// TIA Portal V17 export
// export: Created 2025-07-28T08:20:46.6725827Z, ExportSetting WithDefaults, DisplayName Totally Integrated Automation Portal, DisplayVersion V17, DisplayName TIA Portal Openness, DisplayVersion V17, DisplayName TIA Portal Version Control Interface, DisplayVersion V17, DisplayName SINAMICS Startdrive Advanced, DisplayVersion V17, DisplayName SINAMICS Startdrive G130, G150, S120, S150, SINAMICS MV, S210, DisplayVersion V17, DisplayName SINAMICS Startdrive G110M, G120, G120C, G120D, G120P, G115D, DisplayVersion V17, DisplayName STEP 7 Professional, DisplayVersion V17, DisplayName STEP 7 Safety, DisplayVersion V17, DisplayName WinCC Professional, DisplayVersion V17
FUNCTION_BLOCK "S31808022001_Sequence_All_73b5c5_cfdfd9eb-ebd8-4267-a68e-df0ebcea3fa8 - Copy (2)_f93786"   // FB1, LAD
VERSION : 0.1
// stored: AutoNumber true, IsIECCheckEnabled false, UDAEnableTagReadback false
   VAR_INPUT
      iAutoRunning : Bool;
      iFaultReset : Bool;
      iOTS_Frm_Prev_TTDown : Bool;
      iOTS_Frm_Prev_TTUp : Bool;
      iPalletNtPrsntAtTTDown : Bool;
      iPalletNtPrsntAtTTUp : Bool;
      iPalletPrsnt_TTDown : Bool;
      iPalletPrsnt_TTUp : Bool;
      iPartReject : Bool;
      iRTR_Frm_Next_0DegTTUp : Bool;
      iRTR_Frm_Next_90DegTTUp : Bool;
      iRTR_Frm_Next_TTDown : Bool;
      iRecvAreaClr_TTDown : Bool;
      iRecvAreaClr_TTUp : Bool;
      iReset_fault : Bool;
      iRx_Frm_Prev_TTUp : Bool;
      iSstMode : Bool;
      iSstPB : Bool;
      iStprRaise_TTDown : Bool;
      iStprRaise_TTUp : Bool;
      iTTAt0Pos : Bool;
      iTTAt90Pos : Bool;
      iTTLocked : Bool;
      iTTUnlocked : Bool;
      iXferAreaClr_0DegTTDown : Bool;
      iXferAreaClr_0DegTTUp : Bool;
      iXferAreaClr_90DegTTUp : Bool;
   END_VAR
   VAR_OUTPUT
      qConvRun_TTDown : Bool;
      qConvRun_TTUp : Bool;
      qDelStprDown_TTUp : Bool;
      qOTS_Frm_TTDown : Bool;
      qOTS_Frm_TTUp : Bool;
      qOutput1 : Bool;
      qProcessStart : Bool;
      qRTR_Frm_TTDwn : Bool;
      qRTR_Frm_TTUp : Bool;
      qStprDown_TTDown : Bool;
      qStprDown_TTUp : Bool;
      qStprRaise_TTDown : Bool;
      qStprRaise_TTUp : Bool;
      qTTLockCmd : Bool;
      qTTUnlockCmd : Bool;
      qTT_0Deg : Bool;
      qTT_90Deg : Bool;
   END_VAR
   VAR_IN_OUT
      iqRX_Frn_Prev_TtDown : Bool;
      iqRx_Frm_Prev_TTUp : Bool;
      iqTx_To_Next_0DegTTDown : Bool;
      iqTx_To_Next_0DegTTUp : Bool;
      iqTx_To_Next_90DegTTUp : Bool;
   END_VAR
   VAR DB_SPECIFIC
      StateNo : Int;
      s100_StWtForTTUnlck : Bool;
      s100_StWtForTTUnlck_T1 : Bool;
      s10_StRecoveryCondition : Bool;
      s10_StRecoveryCondition_T1 : Bool;
      s10_StRecoveryCondition_T2 : Bool;
      s10_StRecoveryCondition_T3 : Bool;
      s10_StRecoveryCondition_T4 : Bool;
      s10_StRecoveryCondition_T5 : Bool;
      s10_StRecoveryCondition_T6 : Bool;
      s10_StRecoveryCondition_T7 : Bool;
      s110_StWtForTTTurn90 : Bool;
      s110_StWtForTTTurn90_T1 : Bool;
      s120_StWtForTTLck : Bool;
      s120_StWtForTTLck_T1 : Bool;
      s130_StChkTTDwnRdyToRecv : Bool;
      s130_StChkTTDwnRdyToRecv_T1 : Bool;
      s130_StChkTTDwnRdyToRecv_T2 : Bool;
      s140_StWtFrConveyorStrt : Bool;
      s140_StWtFrConveyorStrt_T1 : Bool;
      s150_StChkNxtStRdyToRecvTTUp : Bool;
      s150_StChkNxtStRdyToRecvTTUp_T1 : Bool;
      s150_StChkNxtStRdyToRecvTTUp_T2 : Bool;
      s15_StWaitForManCorrection : Bool;
      s15_StWaitForManCorrection_T1 : Bool;
      s160_StWtFrStprDn_CnvyrStrt : Bool;
      s160_StWtFrStprDn_CnvyrStrt_T1 : Bool;
      s165_StWtPalAbsnt : Bool;
      s165_StWtPalAbsnt_T1 : Bool;
      s167_StWtFrDeforkOvr : Bool;
      s167_StWtFrDeforkOvr_Cond1 : Bool;
      s167_StWtFrDeforkOvr_Cond2 : Bool;
      s167_StWtFrDeforkOvr_T1 : Bool;
      s170_StWtForTTUpStprUp : Bool;
      s170_StWtForTTUpStprUp_T1 : Bool;
      s180_StWtForTTUnlk : Bool;
      s180_StWtForTTUnlk_T1 : Bool;
      s190_StWtForTT_To_0 : Bool;
      s190_StWtForTT_To_0_T1 : Bool;
      s192_StWtForTTlok : Bool;
      s192_StWtForTTlok_T1 : Bool;
      s20_StChkForPalletPresent : Bool;
      s20_StChkForPalletPresent_T1 : Bool;
      s20_StChkForPalletPresent_T2 : Bool;
      s20_StChkForPalletPresent_T3 : Bool;
      s20_StChkForPalletPresent_T4 : Bool;
      s210_StWtFrTTUnlk : Bool;
      s210_StWtFrTTUnlk_T1 : Bool;
      s220_StWtFrTT_Trn_0 : Bool;
      s220_StWtFrTT_Trn_0_T1 : Bool;
      s230_StWtFrTTLock : Bool;
      s230_StWtFrTTLock_T1 : Bool;
      s240_StWtFRTRNxtStnTTDown : Bool;
      s240_StWtFRTRNxtStnTTDown_T1 : Bool;
      s240_StWtFRTRNxtStnTTDown_T2 : Bool;
      s250_StWtTTDnStprDn_CnvyrStr : Bool;
      s250_StWtTTDnStprDn_CnvyrStr_T1 : Bool;
      s260_StWtPalAbsent : Bool;
      s260_StWtPalAbsent_T1 : Bool;
      s270_StWtFrTTDwnStprUp : Bool;
      s270_StWtFrTTDwnStprUp_T1 : Bool;
      s280_StWtRFrOTSFRmPrev_TTUp : Bool;
      s280_StWtRFrOTSFRmPrev_TTUp_T1 : Bool;
      s290_StWtFrTTUpCnvyrStrt : Bool;
      s290_StWtFrTTUpCnvyrStrt_T1 : Bool;
      s300_StChkTTPos : Bool;
      s300_StChkTTPos_T1 : Bool;
      s300_StChkTTPos_T2 : Bool;
      s300_StChkTTPos_T3 : Bool;
      s30_StChckPartSts : Bool;
      s30_StChckPartSts_T1 : Bool;
      s310_StWtRTRFrmTTUpAt0 : Bool;
      s310_StWtRTRFrmTTUpAt0_T1 : Bool;
      s310_StWtRTRFrmTTUpAt0_T2 : Bool;
      s320_StWtFrTTUpCnvyrStrtAt0 : Bool;
      s320_StWtFrTTUpCnvyrStrtAt0_T1 : Bool;
      s340_StChkTTDwnRdyToRecvAt90 : Bool;
      s340_StChkTTDwnRdyToRecvAt90_T1 : Bool;
      s340_StChkTTDwnRdyToRecvAt90_T2 : Bool;
      s350_StWtCnvyrStrt90 : Bool;
      s350_StWtCnvyrStrt90_T1 : Bool;
      s365_StWtForTTUlkAtIbtwn : Bool;
      s365_StWtForTTUlkAtIbtwn_T1 : Bool;
      s370_StWtForTTTurnZrAtIbtwn : Bool;
      s370_StWtForTTTurnZrAtIbtwn_T1 : Bool;
      s380_StWtForTTLock : Bool;
      s380_StWtForTTLock_T1 : Bool;
      s400_StWt2Defork : Bool;
      s400_StWt2Defork_Cond1 : Bool;
      s400_StWt2Defork_Cond2 : Bool;
      s400_StWt2Defork_T1 : Bool;
      s40_StWtForTTUnlock : Bool;
      s40_StWtForTTUnlock_T1 : Bool;
      s410_StWtForTTUlkAtIbtwn : Bool;
      s410_StWtForTTUlkAtIbtwn_T1 : Bool;
      s415_StWtForTTTurn90AtIbtwn : Bool;
      s415_StWtForTTTurn90AtIbtwn_T1 : Bool;
      s420_StWtForTTLock1 : Bool;
      s420_StWtForTTLock1_T1 : Bool;
      s50_StWtForTTTurn0 : Bool;
      s50_StWtForTTTurn0_T1 : Bool;
      s60_StWtForTTLock : Bool;
      s60_StWtForTTLock_T1 : Bool;
      s70_StWtOTSfrmTTUp : Bool;
      s70_StWtOTSfrmTTUp_T1 : Bool;
      s80_StWtTTUpStpDwnCnvrStrt : Bool;
      s80_StWtTTUpStpDwnCnvrStrt_T1 : Bool;
      s85_StWtPalPresntAtRej : Bool;
      s85_StWtPalPresntAtRej_T1 : Bool;
      s90_StWtTTUpStprUp : Bool;
      s90_StWtTTUpStprUp_T1 : Bool;
      sDefork1Done : Bool;
      sDefork2Done : Bool;
      sOTSFrmDwnTout : Bool;
      sOTSFrmUpTout : Bool;
      sPalOnStop_TTDown : Bool;
      sPalOnStop_TTUp_0Deg : Bool;
      sPalOnStop_TTUp_90Deg : Bool;
      sPalletAbsnDebTTUp : Bool;
      sPalletAbsntDebTTDown : Bool;
      sPalletAbsntDebTTUp : Bool;
      sPalletPrsntDebTTDown : Bool;
      sPalletPrsntDebTTUp : Bool;
      sRTRFrmUpTout : Bool;
      sSst : Bool;
      sSstPulse : Bool;
      sSstRise : Bool;
      sStWtResetRel : Bool;
      sStWtResetRel_T1 : Bool;
      sTTDwnSeqOver : Bool;
      sTTDwn_0Pos_TX_Time : Bool;
      sTTDwn_90Pos_RX_Time : Bool;
      sTTDwn_Timer_ON : Bool;
      sTTUpSeqOver : Bool;
      sTTUp_90Pos_TX_Time : Bool;
      sTTUp_Timer_ON : Bool;
      sTrBothPalletPresent : Bool;
   END_VAR
   VAR_TEMP
      tOne : Bool;
   END_VAR
   VAR_TEMP   // added for the SCL form of the ladder/FBD networks
      _w1 : Bool;
   END_VAR
BEGIN

REGION Network 1
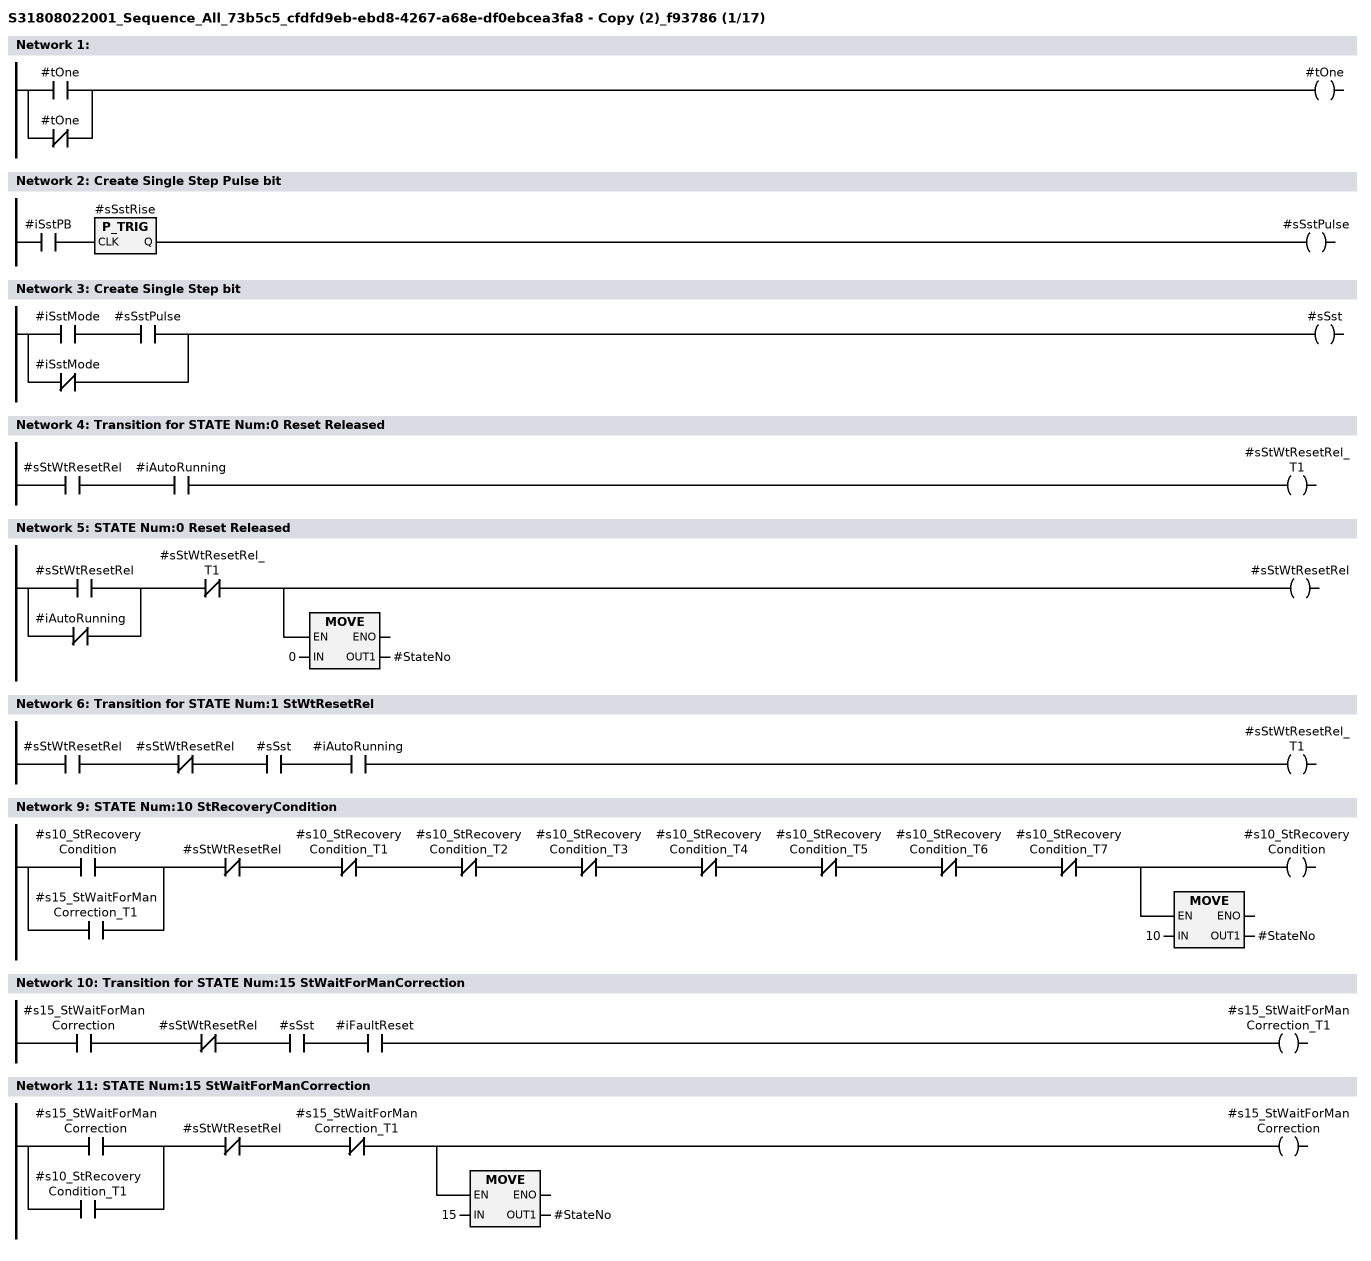
   RUNG wire#powerrail
      Contact( #tOne )
      wire#w1
      Coil( #tOne )
   END_RUNG
   RUNG wire#powerrail
      I_Contact( #tOne )
   END_RUNG wire#w1
   // the same network as SCL:
   #tOne := #tOne OR NOT #tOne;
END_REGION

REGION Network 2: Create Single Step Pulse bit
   RUNG wire#powerrail
      Contact( #iSstPB )
      P_Trig( #sSstRise )
      Coil( #sSstPulse )
   END_RUNG
   // the same network as SCL:
   #_w1 := #iSstPB AND NOT #sSstRise;   // rising edge
   #sSstRise := #iSstPB;
   #sSstPulse := #_w1;
END_REGION

REGION Network 3: Create Single Step bit
   RUNG wire#powerrail
      Contact( #iSstMode )
      Contact( #sSstPulse )
      wire#w1
      Coil( #sSst )
   END_RUNG
   RUNG wire#powerrail
      I_Contact( #iSstMode )
   END_RUNG wire#w1
   // the same network as SCL:
   #sSst := (#iSstMode AND #sSstPulse) OR NOT #iSstMode;
END_REGION

REGION Network 4: Transition for STATE Num:0 Reset Released
   RUNG wire#powerrail
      Contact( #sStWtResetRel )
      Contact( #iAutoRunning )
      Coil( #sStWtResetRel_T1 )
   END_RUNG
   // the same network as SCL:
   #sStWtResetRel_T1 := #sStWtResetRel AND #iAutoRunning;
END_REGION

REGION Network 5: STATE Num:0 Reset Released
   RUNG wire#powerrail
      Contact( #sStWtResetRel )
      wire#w1
      I_Contact( #sStWtResetRel_T1 )
      wire#w2
      Coil( #sStWtResetRel )
   END_RUNG
   RUNG wire#powerrail
      I_Contact( #iAutoRunning )
   END_RUNG wire#w1
   RUNG wire#w2
      { S7_GenerateENO := "TRUE" } Move(in := 0, out1 => #StateNo)
   END_RUNG
   // the same network as SCL:
   #sStWtResetRel := (#sStWtResetRel OR NOT #iAutoRunning) AND NOT #sStWtResetRel_T1;
   IF #sStWtResetRel THEN #StateNo := 0; END_IF;
END_REGION

REGION Network 6: Transition for STATE Num:1 StWtResetRel
   RUNG wire#powerrail
      Contact( #sStWtResetRel )
      I_Contact( #sStWtResetRel )
      Contact( #sSst )
      Contact( #iAutoRunning )
      Coil( #sStWtResetRel_T1 )
   END_RUNG
   // the same network as SCL:
   #sStWtResetRel_T1 := #sStWtResetRel AND NOT #sStWtResetRel AND #sSst AND #iAutoRunning;
END_REGION

NETWORK
TITLE = STATE Num:1 StWtResetRel
      A(;
      O     #sStWtResetRel;
//wrong transition variable removed
      );
      AN    #sStWtResetRel;
      AN    #sStWtResetRel_T1;
      =     %L1.0;
      A     %L1.0;
      BLD   102;
      =     #sStWtResetRel;
      A     %L1.0;
      JNB   Label_1;
      L     1;
      T     #StateNo;
Label_1:NOP   0;

NETWORK
TITLE = Transition for STATE Num:10 StRecoveryCondition
      A     #s10_StRecoveryCondition;
      AN    #sStWtResetRel;
      A     #sSst;
      =     %L1.0;
      A     %L1.0;
      A(;
      O(;
      A     #iRx_Frm_Prev_TTUp;
      AN    #iTTAt0Pos;
      );
      O(;
      A     #iqRX_Frn_Prev_TtDown;
      AN    #iTTAt90Pos;
      );
      O(;
      O     #iqTx_To_Next_90DegTTUp;
      O     #sPalOnStop_TTUp_90Deg;
      AN    #iTTAt90Pos;
      );
      O(;
      O     #iqTx_To_Next_0DegTTUp;
      O     #sPalOnStop_TTUp_0Deg;
      AN    #iTTAt0Pos;
      );
      O(;
      O     #iqTx_To_Next_0DegTTDown;
      O     #sPalOnStop_TTDown;
      AN    #iTTAt0Pos;
      );
      O(;
      O     #sPalOnStop_TTUp_0Deg;
      O     #sPalOnStop_TTUp_90Deg;
      O     #sPalOnStop_TTDown;
      A     #iTTUnlocked;
      );
      );
      =     #s10_StRecoveryCondition_T1;
      A     %L1.0;
      AN    #s10_StRecoveryCondition_T1;
      A(;
      O     #iqTx_To_Next_0DegTTUp;
      O     #sPalOnStop_TTUp_0Deg;
      );
      A     #iTTAt0Pos;
      A     #iTTLocked;
      =     #s10_StRecoveryCondition_T2;
      A     %L1.0;
      AN    #s10_StRecoveryCondition_T1;
      AN    #s10_StRecoveryCondition_T2;
      A(;
      O     #iqTx_To_Next_90DegTTUp;
      O     #sPalOnStop_TTUp_90Deg;
      );
      A     #iTTAt90Pos;
      A     #iTTLocked;
      =     #s10_StRecoveryCondition_T3;
      A     %L1.0;
      AN    #s10_StRecoveryCondition_T1;
      AN    #s10_StRecoveryCondition_T2;
      AN    #s10_StRecoveryCondition_T3;
      A(;
      O     #iqTx_To_Next_0DegTTDown;
      O     #sPalOnStop_TTDown;
      );
      A     #iTTAt0Pos;
      A     #iTTLocked;
      =     #s10_StRecoveryCondition_T4;
      A     %L1.0;
      AN    #s10_StRecoveryCondition_T1;
      AN    #s10_StRecoveryCondition_T2;
      AN    #s10_StRecoveryCondition_T3;
      AN    #s10_StRecoveryCondition_T4;
      A(;
      O     #iRx_Frm_Prev_TTUp;
      O     #iRecvAreaClr_TTUp;
      );
      A     #iTTAt0Pos;
      A     #iTTLocked;
      =     #s10_StRecoveryCondition_T5;
      A     %L1.0;
      AN    #s10_StRecoveryCondition_T1;
      AN    #s10_StRecoveryCondition_T2;
      AN    #s10_StRecoveryCondition_T3;
      AN    #s10_StRecoveryCondition_T4;
      AN    #s10_StRecoveryCondition_T5;
      A(;
      O     #iqRX_Frn_Prev_TtDown;
      ON    #iRecvAreaClr_TTDown;
      );
      A     #iTTAt90Pos;
      A     #iTTLocked;
      =     #s10_StRecoveryCondition_T6;
      A     %L1.0;
      AN    #s10_StRecoveryCondition_T1;
      AN    #s10_StRecoveryCondition_T2;
      AN    #s10_StRecoveryCondition_T3;
      AN    #s10_StRecoveryCondition_T4;
      AN    #s10_StRecoveryCondition_T5;
      AN    #s10_StRecoveryCondition_T6;
      A(;
      A(;
      A     #iXferAreaClr_90DegTTUp;
      A     #iXferAreaClr_0DegTTDown;
      A     #iRecvAreaClr_TTDown;
      A     #iRecvAreaClr_TTUp;
      );
      O(;
      AN    #sPalOnStop_TTUp_0Deg;
      AN    #sPalOnStop_TTUp_90Deg;
      AN    #sPalOnStop_TTDown;
      );
      O(;
      AN    #iqTx_To_Next_90DegTTUp;
      AN    #iqTx_To_Next_0DegTTUp;
      AN    #iqTx_To_Next_0DegTTDown;
      AN    #iqRX_Frn_Prev_TtDown;
      AN    #iRx_Frm_Prev_TTUp;
      );
      );
      =     #s10_StRecoveryCondition_T7;

REGION Network 9: STATE Num:10 StRecoveryCondition
   RUNG wire#powerrail
      Contact( #s10_StRecoveryCondition )
      wire#w1
      I_Contact( #sStWtResetRel )
      I_Contact( #s10_StRecoveryCondition_T1 )
      I_Contact( #s10_StRecoveryCondition_T2 )
      I_Contact( #s10_StRecoveryCondition_T3 )
      I_Contact( #s10_StRecoveryCondition_T4 )
      I_Contact( #s10_StRecoveryCondition_T5 )
      I_Contact( #s10_StRecoveryCondition_T6 )
      I_Contact( #s10_StRecoveryCondition_T7 )
      wire#w2
      Coil( #s10_StRecoveryCondition )
   END_RUNG
   RUNG wire#powerrail
      Contact( #s15_StWaitForManCorrection_T1 )
   END_RUNG wire#w1
   RUNG wire#w2
      { S7_GenerateENO := "TRUE" } Move(in := 10, out1 => #StateNo)
   END_RUNG
   // the same network as SCL:
   #s10_StRecoveryCondition := (#s10_StRecoveryCondition OR #s15_StWaitForManCorrection_T1) AND NOT #sStWtResetRel AND NOT #s10_StRecoveryCondition_T1 AND NOT #s10_StRecoveryCondition_T2 AND NOT #s10_StRecoveryCondition_T3 AND NOT #s10_StRecoveryCondition_T4 AND NOT #s10_StRecoveryCondition_T5 AND NOT #s10_StRecoveryCondition_T6 AND NOT #s10_StRecoveryCondition_T7;
   IF #s10_StRecoveryCondition THEN #StateNo := 10; END_IF;
END_REGION

REGION Network 10: Transition for STATE Num:15 StWaitForManCorrection
   RUNG wire#powerrail
      Contact( #s15_StWaitForManCorrection )
      I_Contact( #sStWtResetRel )
      Contact( #sSst )
      Contact( #iFaultReset )
      Coil( #s15_StWaitForManCorrection_T1 )
   END_RUNG
   // the same network as SCL:
   #s15_StWaitForManCorrection_T1 := #s15_StWaitForManCorrection AND NOT #sStWtResetRel AND #sSst AND #iFaultReset;
END_REGION

REGION Network 11: STATE Num:15 StWaitForManCorrection
   RUNG wire#powerrail
      Contact( #s15_StWaitForManCorrection )
      wire#w1
      I_Contact( #sStWtResetRel )
      I_Contact( #s15_StWaitForManCorrection_T1 )
      wire#w2
      Coil( #s15_StWaitForManCorrection )
   END_RUNG
   RUNG wire#powerrail
      Contact( #s10_StRecoveryCondition_T1 )
   END_RUNG wire#w1
   RUNG wire#w2
      { S7_GenerateENO := "TRUE" } Move(in := 15, out1 => #StateNo)
   END_RUNG
   // the same network as SCL:
   #s15_StWaitForManCorrection := (#s15_StWaitForManCorrection OR #s10_StRecoveryCondition_T1) AND NOT #sStWtResetRel AND NOT #s15_StWaitForManCorrection_T1;
   IF #s15_StWaitForManCorrection THEN #StateNo := 15; END_IF;
END_REGION

REGION Network 12: Transition for STATE Num:20 StChkForPalletPresent
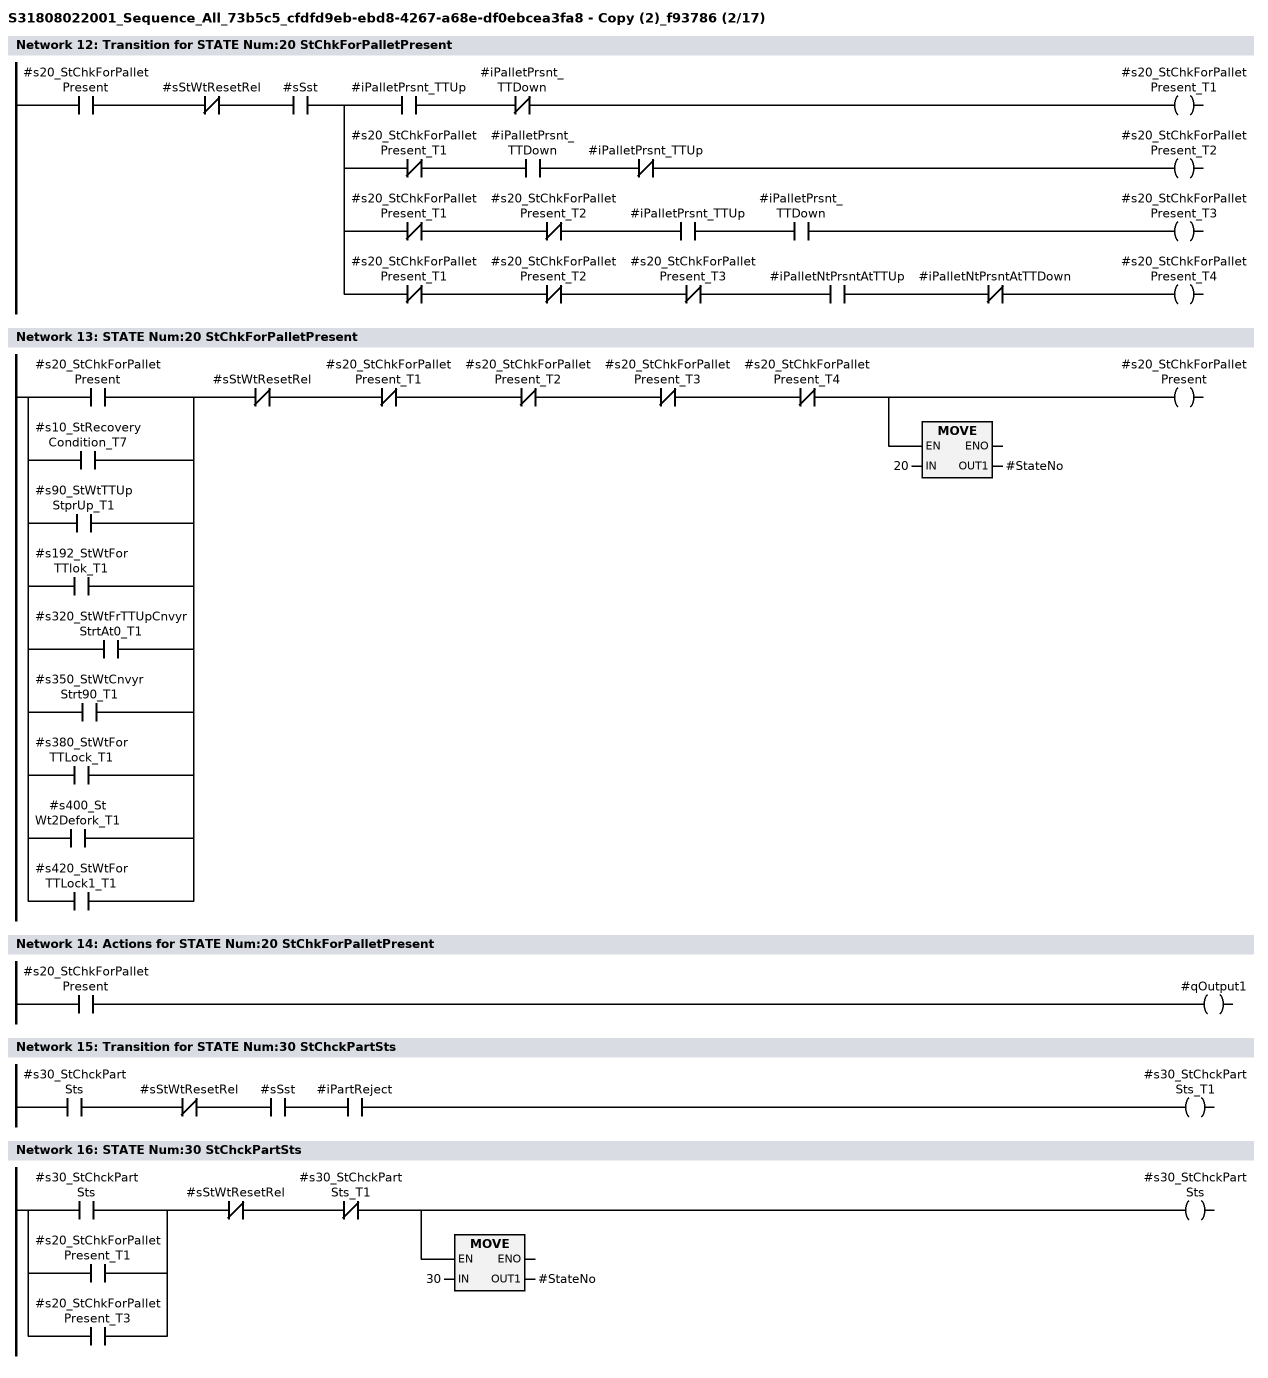
   RUNG wire#powerrail
      Contact( #s20_StChkForPalletPresent )
      I_Contact( #sStWtResetRel )
      Contact( #sSst )
      wire#w1
      Contact( #iPalletPrsnt_TTUp )
      I_Contact( #iPalletPrsnt_TTDown )
      Coil( #s20_StChkForPalletPresent_T1 )
   END_RUNG
   RUNG wire#w1
      I_Contact( #s20_StChkForPalletPresent_T1 )
      Contact( #iPalletPrsnt_TTDown )
      I_Contact( #iPalletPrsnt_TTUp )
      Coil( #s20_StChkForPalletPresent_T2 )
   END_RUNG
   RUNG wire#w1
      I_Contact( #s20_StChkForPalletPresent_T1 )
      I_Contact( #s20_StChkForPalletPresent_T2 )
      Contact( #iPalletPrsnt_TTUp )
      Contact( #iPalletPrsnt_TTDown )
      Coil( #s20_StChkForPalletPresent_T3 )
   END_RUNG
   RUNG wire#w1
      I_Contact( #s20_StChkForPalletPresent_T1 )
      I_Contact( #s20_StChkForPalletPresent_T2 )
      I_Contact( #s20_StChkForPalletPresent_T3 )
      Contact( #iPalletNtPrsntAtTTUp )
      I_Contact( #iPalletNtPrsntAtTTDown )
      Coil( #s20_StChkForPalletPresent_T4 )
   END_RUNG
   // the same network as SCL:
   #_w1 := #s20_StChkForPalletPresent AND NOT #sStWtResetRel AND #sSst;
   #s20_StChkForPalletPresent_T1 := #_w1 AND #iPalletPrsnt_TTUp AND NOT #iPalletPrsnt_TTDown;
   #s20_StChkForPalletPresent_T2 := #_w1 AND NOT #s20_StChkForPalletPresent_T1 AND #iPalletPrsnt_TTDown AND NOT #iPalletPrsnt_TTUp;
   #s20_StChkForPalletPresent_T3 := #_w1 AND NOT #s20_StChkForPalletPresent_T1 AND NOT #s20_StChkForPalletPresent_T2 AND #iPalletPrsnt_TTUp AND #iPalletPrsnt_TTDown;
   #s20_StChkForPalletPresent_T4 := #_w1 AND NOT #s20_StChkForPalletPresent_T1 AND NOT #s20_StChkForPalletPresent_T2 AND NOT #s20_StChkForPalletPresent_T3 AND #iPalletNtPrsntAtTTUp AND NOT #iPalletNtPrsntAtTTDown;
END_REGION

REGION Network 13: STATE Num:20 StChkForPalletPresent
   RUNG wire#powerrail
      Contact( #s20_StChkForPalletPresent )
      wire#w1
      I_Contact( #sStWtResetRel )
      I_Contact( #s20_StChkForPalletPresent_T1 )
      I_Contact( #s20_StChkForPalletPresent_T2 )
      I_Contact( #s20_StChkForPalletPresent_T3 )
      I_Contact( #s20_StChkForPalletPresent_T4 )
      wire#w2
      Coil( #s20_StChkForPalletPresent )
   END_RUNG
   RUNG wire#powerrail
      Contact( #s10_StRecoveryCondition_T7 )
   END_RUNG wire#w1
   RUNG wire#powerrail
      Contact( #s90_StWtTTUpStprUp_T1 )
   END_RUNG wire#w1
   RUNG wire#powerrail
      Contact( #s192_StWtForTTlok_T1 )
   END_RUNG wire#w1
   RUNG wire#powerrail
      Contact( #s320_StWtFrTTUpCnvyrStrtAt0_T1 )
   END_RUNG wire#w1
   RUNG wire#powerrail
      Contact( #s350_StWtCnvyrStrt90_T1 )
   END_RUNG wire#w1
   RUNG wire#powerrail
      Contact( #s380_StWtForTTLock_T1 )
   END_RUNG wire#w1
   RUNG wire#powerrail
      Contact( #s400_StWt2Defork_T1 )
   END_RUNG wire#w1
   RUNG wire#powerrail
      Contact( #s420_StWtForTTLock1_T1 )
   END_RUNG wire#w1
   RUNG wire#w2
      { S7_GenerateENO := "TRUE" } Move(in := 20, out1 => #StateNo)
   END_RUNG
   // the same network as SCL:
   #s20_StChkForPalletPresent := (#s20_StChkForPalletPresent OR #s10_StRecoveryCondition_T7 OR #s90_StWtTTUpStprUp_T1 OR #s192_StWtForTTlok_T1 OR #s320_StWtFrTTUpCnvyrStrtAt0_T1 OR #s350_StWtCnvyrStrt90_T1 OR #s380_StWtForTTLock_T1 OR #s400_StWt2Defork_T1 OR #s420_StWtForTTLock1_T1) AND NOT #sStWtResetRel AND NOT #s20_StChkForPalletPresent_T1 AND NOT #s20_StChkForPalletPresent_T2 AND NOT #s20_StChkForPalletPresent_T3 AND NOT #s20_StChkForPalletPresent_T4;
   IF #s20_StChkForPalletPresent THEN #StateNo := 20; END_IF;
END_REGION

REGION Network 14: Actions for STATE Num:20 StChkForPalletPresent
   RUNG wire#powerrail
      Contact( #s20_StChkForPalletPresent )
      Coil( #qOutput1 )
   END_RUNG
   // the same network as SCL:
   #qOutput1 := #s20_StChkForPalletPresent;
END_REGION

REGION Network 15: Transition for STATE Num:30 StChckPartSts
   RUNG wire#powerrail
      Contact( #s30_StChckPartSts )
      I_Contact( #sStWtResetRel )
      Contact( #sSst )
      Contact( #iPartReject )
      Coil( #s30_StChckPartSts_T1 )
   END_RUNG
   // the same network as SCL:
   #s30_StChckPartSts_T1 := #s30_StChckPartSts AND NOT #sStWtResetRel AND #sSst AND #iPartReject;
END_REGION

REGION Network 16: STATE Num:30 StChckPartSts
   RUNG wire#powerrail
      Contact( #s30_StChckPartSts )
      wire#w1
      I_Contact( #sStWtResetRel )
      I_Contact( #s30_StChckPartSts_T1 )
      wire#w2
      Coil( #s30_StChckPartSts )
   END_RUNG
   RUNG wire#powerrail
      Contact( #s20_StChkForPalletPresent_T1 )
   END_RUNG wire#w1
   RUNG wire#powerrail
      Contact( #s20_StChkForPalletPresent_T3 )
   END_RUNG wire#w1
   RUNG wire#w2
      { S7_GenerateENO := "TRUE" } Move(in := 30, out1 => #StateNo)
   END_RUNG
   // the same network as SCL:
   #s30_StChckPartSts := (#s30_StChckPartSts OR #s20_StChkForPalletPresent_T1 OR #s20_StChkForPalletPresent_T3) AND NOT #sStWtResetRel AND NOT #s30_StChckPartSts_T1;
   IF #s30_StChckPartSts THEN #StateNo := 30; END_IF;
END_REGION

REGION Network 17: Actions for STATE Num:30 StChckPartSts
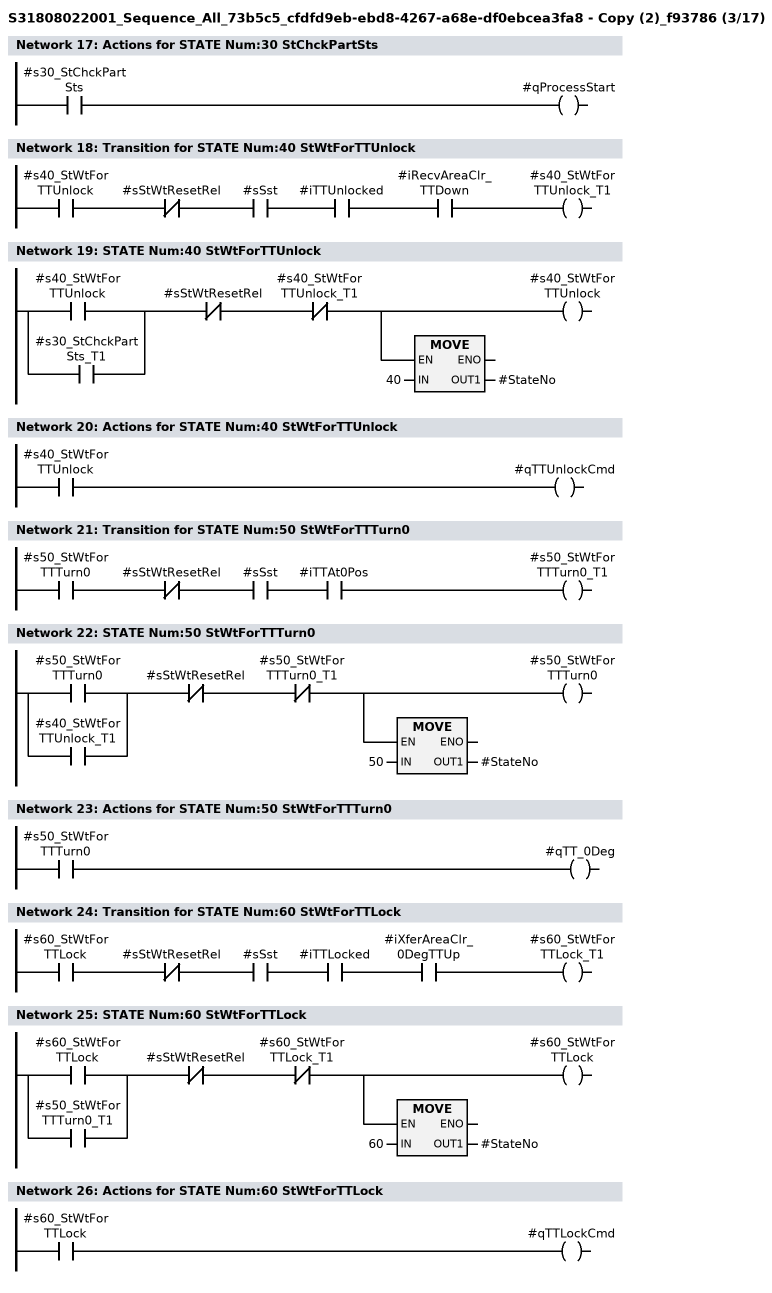
   RUNG wire#powerrail
      Contact( #s30_StChckPartSts )
      Coil( #qProcessStart )
   END_RUNG
   // the same network as SCL:
   #qProcessStart := #s30_StChckPartSts;
END_REGION

REGION Network 18: Transition for STATE Num:40 StWtForTTUnlock
   RUNG wire#powerrail
      Contact( #s40_StWtForTTUnlock )
      I_Contact( #sStWtResetRel )
      Contact( #sSst )
      Contact( #iTTUnlocked )
      Contact( #iRecvAreaClr_TTDown )
      Coil( #s40_StWtForTTUnlock_T1 )
   END_RUNG
   // the same network as SCL:
   #s40_StWtForTTUnlock_T1 := #s40_StWtForTTUnlock AND NOT #sStWtResetRel AND #sSst AND #iTTUnlocked AND #iRecvAreaClr_TTDown;
END_REGION

REGION Network 19: STATE Num:40 StWtForTTUnlock
   RUNG wire#powerrail
      Contact( #s40_StWtForTTUnlock )
      wire#w1
      I_Contact( #sStWtResetRel )
      I_Contact( #s40_StWtForTTUnlock_T1 )
      wire#w2
      Coil( #s40_StWtForTTUnlock )
   END_RUNG
   RUNG wire#powerrail
      Contact( #s30_StChckPartSts_T1 )
   END_RUNG wire#w1
   RUNG wire#w2
      { S7_GenerateENO := "TRUE" } Move(in := 40, out1 => #StateNo)
   END_RUNG
   // the same network as SCL:
   #s40_StWtForTTUnlock := (#s40_StWtForTTUnlock OR #s30_StChckPartSts_T1) AND NOT #sStWtResetRel AND NOT #s40_StWtForTTUnlock_T1;
   IF #s40_StWtForTTUnlock THEN #StateNo := 40; END_IF;
END_REGION

REGION Network 20: Actions for STATE Num:40 StWtForTTUnlock
   RUNG wire#powerrail
      Contact( #s40_StWtForTTUnlock )
      Coil( #qTTUnlockCmd )
   END_RUNG
   // the same network as SCL:
   #qTTUnlockCmd := #s40_StWtForTTUnlock;
END_REGION

REGION Network 21: Transition for STATE Num:50 StWtForTTTurn0
   RUNG wire#powerrail
      Contact( #s50_StWtForTTTurn0 )
      I_Contact( #sStWtResetRel )
      Contact( #sSst )
      Contact( #iTTAt0Pos )
      Coil( #s50_StWtForTTTurn0_T1 )
   END_RUNG
   // the same network as SCL:
   #s50_StWtForTTTurn0_T1 := #s50_StWtForTTTurn0 AND NOT #sStWtResetRel AND #sSst AND #iTTAt0Pos;
END_REGION

REGION Network 22: STATE Num:50 StWtForTTTurn0
   RUNG wire#powerrail
      Contact( #s50_StWtForTTTurn0 )
      wire#w1
      I_Contact( #sStWtResetRel )
      I_Contact( #s50_StWtForTTTurn0_T1 )
      wire#w2
      Coil( #s50_StWtForTTTurn0 )
   END_RUNG
   RUNG wire#powerrail
      Contact( #s40_StWtForTTUnlock_T1 )
   END_RUNG wire#w1
   RUNG wire#w2
      { S7_GenerateENO := "TRUE" } Move(in := 50, out1 => #StateNo)
   END_RUNG
   // the same network as SCL:
   #s50_StWtForTTTurn0 := (#s50_StWtForTTTurn0 OR #s40_StWtForTTUnlock_T1) AND NOT #sStWtResetRel AND NOT #s50_StWtForTTTurn0_T1;
   IF #s50_StWtForTTTurn0 THEN #StateNo := 50; END_IF;
END_REGION

REGION Network 23: Actions for STATE Num:50 StWtForTTTurn0
   RUNG wire#powerrail
      Contact( #s50_StWtForTTTurn0 )
      Coil( #qTT_0Deg )
   END_RUNG
   // the same network as SCL:
   #qTT_0Deg := #s50_StWtForTTTurn0;
END_REGION

REGION Network 24: Transition for STATE Num:60 StWtForTTLock
   RUNG wire#powerrail
      Contact( #s60_StWtForTTLock )
      I_Contact( #sStWtResetRel )
      Contact( #sSst )
      Contact( #iTTLocked )
      Contact( #iXferAreaClr_0DegTTUp )
      Coil( #s60_StWtForTTLock_T1 )
   END_RUNG
   // the same network as SCL:
   #s60_StWtForTTLock_T1 := #s60_StWtForTTLock AND NOT #sStWtResetRel AND #sSst AND #iTTLocked AND #iXferAreaClr_0DegTTUp;
END_REGION

REGION Network 25: STATE Num:60 StWtForTTLock
   RUNG wire#powerrail
      Contact( #s60_StWtForTTLock )
      wire#w1
      I_Contact( #sStWtResetRel )
      I_Contact( #s60_StWtForTTLock_T1 )
      wire#w2
      Coil( #s60_StWtForTTLock )
   END_RUNG
   RUNG wire#powerrail
      Contact( #s50_StWtForTTTurn0_T1 )
   END_RUNG wire#w1
   RUNG wire#w2
      { S7_GenerateENO := "TRUE" } Move(in := 60, out1 => #StateNo)
   END_RUNG
   // the same network as SCL:
   #s60_StWtForTTLock := (#s60_StWtForTTLock OR #s50_StWtForTTTurn0_T1) AND NOT #sStWtResetRel AND NOT #s60_StWtForTTLock_T1;
   IF #s60_StWtForTTLock THEN #StateNo := 60; END_IF;
END_REGION

REGION Network 26: Actions for STATE Num:60 StWtForTTLock
   RUNG wire#powerrail
      Contact( #s60_StWtForTTLock )
      Coil( #qTTLockCmd )
   END_RUNG
   // the same network as SCL:
   #qTTLockCmd := #s60_StWtForTTLock;
END_REGION

REGION Network 27: Transition for STATE Num:70 StWtOTSfrmTTUp
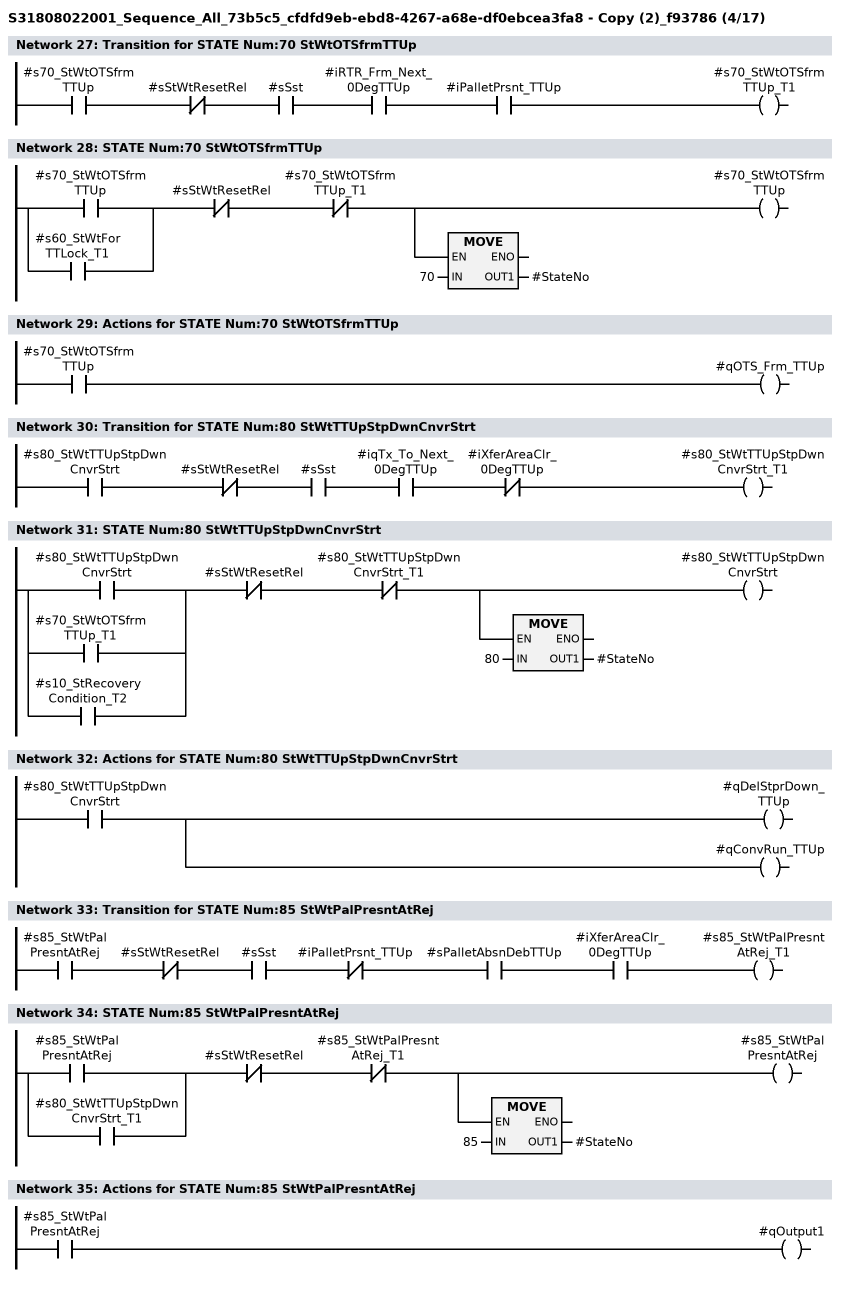
   RUNG wire#powerrail
      Contact( #s70_StWtOTSfrmTTUp )
      I_Contact( #sStWtResetRel )
      Contact( #sSst )
      Contact( #iRTR_Frm_Next_0DegTTUp )
      Contact( #iPalletPrsnt_TTUp )
      Coil( #s70_StWtOTSfrmTTUp_T1 )
   END_RUNG
   // the same network as SCL:
   #s70_StWtOTSfrmTTUp_T1 := #s70_StWtOTSfrmTTUp AND NOT #sStWtResetRel AND #sSst AND #iRTR_Frm_Next_0DegTTUp AND #iPalletPrsnt_TTUp;
END_REGION

REGION Network 28: STATE Num:70 StWtOTSfrmTTUp
   RUNG wire#powerrail
      Contact( #s70_StWtOTSfrmTTUp )
      wire#w1
      I_Contact( #sStWtResetRel )
      I_Contact( #s70_StWtOTSfrmTTUp_T1 )
      wire#w2
      Coil( #s70_StWtOTSfrmTTUp )
   END_RUNG
   RUNG wire#powerrail
      Contact( #s60_StWtForTTLock_T1 )
   END_RUNG wire#w1
   RUNG wire#w2
      { S7_GenerateENO := "TRUE" } Move(in := 70, out1 => #StateNo)
   END_RUNG
   // the same network as SCL:
   #s70_StWtOTSfrmTTUp := (#s70_StWtOTSfrmTTUp OR #s60_StWtForTTLock_T1) AND NOT #sStWtResetRel AND NOT #s70_StWtOTSfrmTTUp_T1;
   IF #s70_StWtOTSfrmTTUp THEN #StateNo := 70; END_IF;
END_REGION

REGION Network 29: Actions for STATE Num:70 StWtOTSfrmTTUp
   RUNG wire#powerrail
      Contact( #s70_StWtOTSfrmTTUp )
      Coil( #qOTS_Frm_TTUp )
   END_RUNG
   // the same network as SCL:
   #qOTS_Frm_TTUp := #s70_StWtOTSfrmTTUp;
END_REGION

REGION Network 30: Transition for STATE Num:80 StWtTTUpStpDwnCnvrStrt
   RUNG wire#powerrail
      Contact( #s80_StWtTTUpStpDwnCnvrStrt )
      I_Contact( #sStWtResetRel )
      Contact( #sSst )
      Contact( #iqTx_To_Next_0DegTTUp )
      I_Contact( #iXferAreaClr_0DegTTUp )
      Coil( #s80_StWtTTUpStpDwnCnvrStrt_T1 )
   END_RUNG
   // the same network as SCL:
   #s80_StWtTTUpStpDwnCnvrStrt_T1 := #s80_StWtTTUpStpDwnCnvrStrt AND NOT #sStWtResetRel AND #sSst AND #iqTx_To_Next_0DegTTUp AND NOT #iXferAreaClr_0DegTTUp;
END_REGION

REGION Network 31: STATE Num:80 StWtTTUpStpDwnCnvrStrt
   RUNG wire#powerrail
      Contact( #s80_StWtTTUpStpDwnCnvrStrt )
      wire#w1
      I_Contact( #sStWtResetRel )
      I_Contact( #s80_StWtTTUpStpDwnCnvrStrt_T1 )
      wire#w2
      Coil( #s80_StWtTTUpStpDwnCnvrStrt )
   END_RUNG
   RUNG wire#powerrail
      Contact( #s70_StWtOTSfrmTTUp_T1 )
   END_RUNG wire#w1
   RUNG wire#powerrail
      Contact( #s10_StRecoveryCondition_T2 )
   END_RUNG wire#w1
   RUNG wire#w2
      { S7_GenerateENO := "TRUE" } Move(in := 80, out1 => #StateNo)
   END_RUNG
   // the same network as SCL:
   #s80_StWtTTUpStpDwnCnvrStrt := (#s80_StWtTTUpStpDwnCnvrStrt OR #s70_StWtOTSfrmTTUp_T1 OR #s10_StRecoveryCondition_T2) AND NOT #sStWtResetRel AND NOT #s80_StWtTTUpStpDwnCnvrStrt_T1;
   IF #s80_StWtTTUpStpDwnCnvrStrt THEN #StateNo := 80; END_IF;
END_REGION

REGION Network 32: Actions for STATE Num:80 StWtTTUpStpDwnCnvrStrt
   RUNG wire#powerrail
      Contact( #s80_StWtTTUpStpDwnCnvrStrt )
      wire#w1
      Coil( #qDelStprDown_TTUp )
   END_RUNG
   RUNG wire#w1
      Coil( #qConvRun_TTUp )
   END_RUNG
   // the same network as SCL:
   #qDelStprDown_TTUp := #s80_StWtTTUpStpDwnCnvrStrt;
   #qConvRun_TTUp := #s80_StWtTTUpStpDwnCnvrStrt;
END_REGION

REGION Network 33: Transition for STATE Num:85 StWtPalPresntAtRej
   RUNG wire#powerrail
      Contact( #s85_StWtPalPresntAtRej )
      I_Contact( #sStWtResetRel )
      Contact( #sSst )
      I_Contact( #iPalletPrsnt_TTUp )
      Contact( #sPalletAbsnDebTTUp )
      Contact( #iXferAreaClr_0DegTTUp )
      Coil( #s85_StWtPalPresntAtRej_T1 )
   END_RUNG
   // the same network as SCL:
   #s85_StWtPalPresntAtRej_T1 := #s85_StWtPalPresntAtRej AND NOT #sStWtResetRel AND #sSst AND NOT #iPalletPrsnt_TTUp AND #sPalletAbsnDebTTUp AND #iXferAreaClr_0DegTTUp;
END_REGION

REGION Network 34: STATE Num:85 StWtPalPresntAtRej
   RUNG wire#powerrail
      Contact( #s85_StWtPalPresntAtRej )
      wire#w1
      I_Contact( #sStWtResetRel )
      I_Contact( #s85_StWtPalPresntAtRej_T1 )
      wire#w2
      Coil( #s85_StWtPalPresntAtRej )
   END_RUNG
   RUNG wire#powerrail
      Contact( #s80_StWtTTUpStpDwnCnvrStrt_T1 )
   END_RUNG wire#w1
   RUNG wire#w2
      { S7_GenerateENO := "TRUE" } Move(in := 85, out1 => #StateNo)
   END_RUNG
   // the same network as SCL:
   #s85_StWtPalPresntAtRej := (#s85_StWtPalPresntAtRej OR #s80_StWtTTUpStpDwnCnvrStrt_T1) AND NOT #sStWtResetRel AND NOT #s85_StWtPalPresntAtRej_T1;
   IF #s85_StWtPalPresntAtRej THEN #StateNo := 85; END_IF;
END_REGION

REGION Network 35: Actions for STATE Num:85 StWtPalPresntAtRej
   RUNG wire#powerrail
      Contact( #s85_StWtPalPresntAtRej )
      Coil( #qOutput1 )
   END_RUNG
   // the same network as SCL:
   #qOutput1 := #s85_StWtPalPresntAtRej;
END_REGION

REGION Network 36: Transition for STATE Num:90 StWtTTUpStprUp
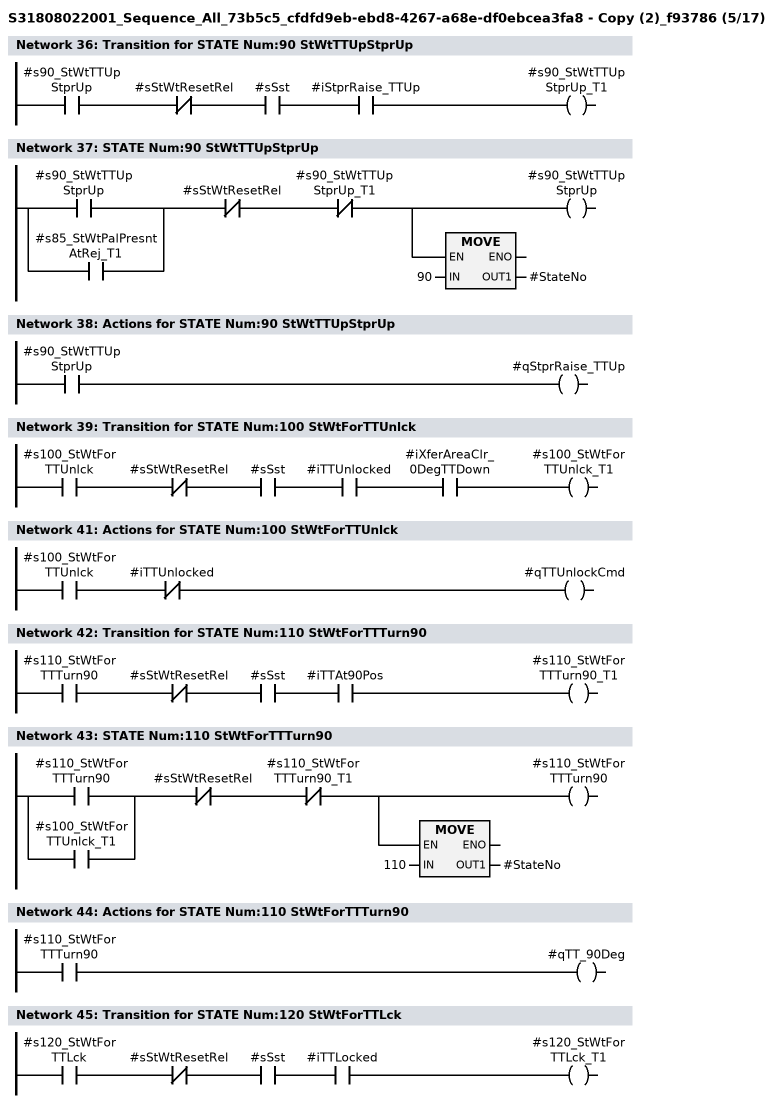
   RUNG wire#powerrail
      Contact( #s90_StWtTTUpStprUp )
      I_Contact( #sStWtResetRel )
      Contact( #sSst )
      Contact( #iStprRaise_TTUp )
      Coil( #s90_StWtTTUpStprUp_T1 )
   END_RUNG
   // the same network as SCL:
   #s90_StWtTTUpStprUp_T1 := #s90_StWtTTUpStprUp AND NOT #sStWtResetRel AND #sSst AND #iStprRaise_TTUp;
END_REGION

REGION Network 37: STATE Num:90 StWtTTUpStprUp
   RUNG wire#powerrail
      Contact( #s90_StWtTTUpStprUp )
      wire#w1
      I_Contact( #sStWtResetRel )
      I_Contact( #s90_StWtTTUpStprUp_T1 )
      wire#w2
      Coil( #s90_StWtTTUpStprUp )
   END_RUNG
   RUNG wire#powerrail
      Contact( #s85_StWtPalPresntAtRej_T1 )
   END_RUNG wire#w1
   RUNG wire#w2
      { S7_GenerateENO := "TRUE" } Move(in := 90, out1 => #StateNo)
   END_RUNG
   // the same network as SCL:
   #s90_StWtTTUpStprUp := (#s90_StWtTTUpStprUp OR #s85_StWtPalPresntAtRej_T1) AND NOT #sStWtResetRel AND NOT #s90_StWtTTUpStprUp_T1;
   IF #s90_StWtTTUpStprUp THEN #StateNo := 90; END_IF;
END_REGION

REGION Network 38: Actions for STATE Num:90 StWtTTUpStprUp
   RUNG wire#powerrail
      Contact( #s90_StWtTTUpStprUp )
      Coil( #qStprRaise_TTUp )
   END_RUNG
   // the same network as SCL:
   #qStprRaise_TTUp := #s90_StWtTTUpStprUp;
END_REGION

REGION Network 39: Transition for STATE Num:100 StWtForTTUnlck
   RUNG wire#powerrail
      Contact( #s100_StWtForTTUnlck )
      I_Contact( #sStWtResetRel )
      Contact( #sSst )
      Contact( #iTTUnlocked )
      Contact( #iXferAreaClr_0DegTTDown )
      Coil( #s100_StWtForTTUnlck_T1 )
   END_RUNG
   // the same network as SCL:
   #s100_StWtForTTUnlck_T1 := #s100_StWtForTTUnlck AND NOT #sStWtResetRel AND #sSst AND #iTTUnlocked AND #iXferAreaClr_0DegTTDown;
END_REGION

NETWORK
TITLE = STATE Num:100 StWtForTTUnlck
      A(;
      O     #s100_StWtForTTUnlck;
      );
      AN    #sStWtResetRel;
      AN    #s100_StWtForTTUnlck_T1;
      =     %L1.0;
      A     %L1.0;
      BLD   102;
      =     #s100_StWtForTTUnlck;
      A     %L1.0;
      JNB   Label_13;
      L     100;
      T     #StateNo;
Label_13:NOP   0;

REGION Network 41: Actions for STATE Num:100 StWtForTTUnlck
   RUNG wire#powerrail
      Contact( #s100_StWtForTTUnlck )
      I_Contact( #iTTUnlocked )
      Coil( #qTTUnlockCmd )
   END_RUNG
   // the same network as SCL:
   #qTTUnlockCmd := #s100_StWtForTTUnlck AND NOT #iTTUnlocked;
END_REGION

REGION Network 42: Transition for STATE Num:110 StWtForTTTurn90
   RUNG wire#powerrail
      Contact( #s110_StWtForTTTurn90 )
      I_Contact( #sStWtResetRel )
      Contact( #sSst )
      Contact( #iTTAt90Pos )
      Coil( #s110_StWtForTTTurn90_T1 )
   END_RUNG
   // the same network as SCL:
   #s110_StWtForTTTurn90_T1 := #s110_StWtForTTTurn90 AND NOT #sStWtResetRel AND #sSst AND #iTTAt90Pos;
END_REGION

REGION Network 43: STATE Num:110 StWtForTTTurn90
   RUNG wire#powerrail
      Contact( #s110_StWtForTTTurn90 )
      wire#w1
      I_Contact( #sStWtResetRel )
      I_Contact( #s110_StWtForTTTurn90_T1 )
      wire#w2
      Coil( #s110_StWtForTTTurn90 )
   END_RUNG
   RUNG wire#powerrail
      Contact( #s100_StWtForTTUnlck_T1 )
   END_RUNG wire#w1
   RUNG wire#w2
      { S7_GenerateENO := "TRUE" } Move(in := 110, out1 => #StateNo)
   END_RUNG
   // the same network as SCL:
   #s110_StWtForTTTurn90 := (#s110_StWtForTTTurn90 OR #s100_StWtForTTUnlck_T1) AND NOT #sStWtResetRel AND NOT #s110_StWtForTTTurn90_T1;
   IF #s110_StWtForTTTurn90 THEN #StateNo := 110; END_IF;
END_REGION

REGION Network 44: Actions for STATE Num:110 StWtForTTTurn90
   RUNG wire#powerrail
      Contact( #s110_StWtForTTTurn90 )
      Coil( #qTT_90Deg )
   END_RUNG
   // the same network as SCL:
   #qTT_90Deg := #s110_StWtForTTTurn90;
END_REGION

REGION Network 45: Transition for STATE Num:120 StWtForTTLck
   RUNG wire#powerrail
      Contact( #s120_StWtForTTLck )
      I_Contact( #sStWtResetRel )
      Contact( #sSst )
      Contact( #iTTLocked )
      Coil( #s120_StWtForTTLck_T1 )
   END_RUNG
   // the same network as SCL:
   #s120_StWtForTTLck_T1 := #s120_StWtForTTLck AND NOT #sStWtResetRel AND #sSst AND #iTTLocked;
END_REGION

REGION Network 46: STATE Num:120 StWtForTTLck
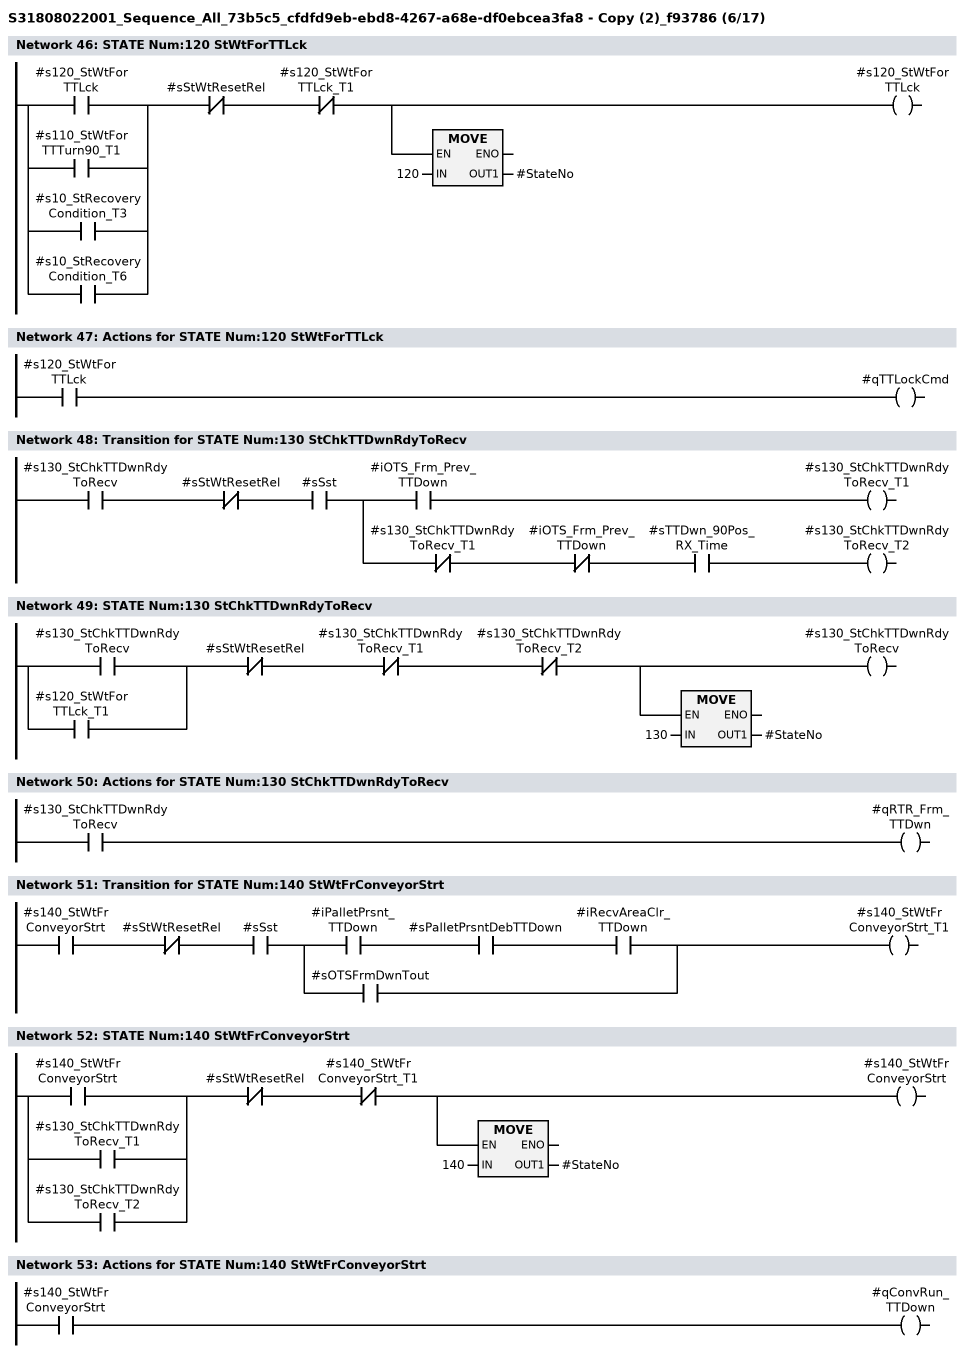
   RUNG wire#powerrail
      Contact( #s120_StWtForTTLck )
      wire#w1
      I_Contact( #sStWtResetRel )
      I_Contact( #s120_StWtForTTLck_T1 )
      wire#w2
      Coil( #s120_StWtForTTLck )
   END_RUNG
   RUNG wire#powerrail
      Contact( #s110_StWtForTTTurn90_T1 )
   END_RUNG wire#w1
   RUNG wire#powerrail
      Contact( #s10_StRecoveryCondition_T3 )
   END_RUNG wire#w1
   RUNG wire#powerrail
      Contact( #s10_StRecoveryCondition_T6 )
   END_RUNG wire#w1
   RUNG wire#w2
      { S7_GenerateENO := "TRUE" } Move(in := 120, out1 => #StateNo)
   END_RUNG
   // the same network as SCL:
   #s120_StWtForTTLck := (#s120_StWtForTTLck OR #s110_StWtForTTTurn90_T1 OR #s10_StRecoveryCondition_T3 OR #s10_StRecoveryCondition_T6) AND NOT #sStWtResetRel AND NOT #s120_StWtForTTLck_T1;
   IF #s120_StWtForTTLck THEN #StateNo := 120; END_IF;
END_REGION

REGION Network 47: Actions for STATE Num:120 StWtForTTLck
   RUNG wire#powerrail
      Contact( #s120_StWtForTTLck )
      Coil( #qTTLockCmd )
   END_RUNG
   // the same network as SCL:
   #qTTLockCmd := #s120_StWtForTTLck;
END_REGION

REGION Network 48: Transition for STATE Num:130 StChkTTDwnRdyToRecv
   RUNG wire#powerrail
      Contact( #s130_StChkTTDwnRdyToRecv )
      I_Contact( #sStWtResetRel )
      Contact( #sSst )
      wire#w1
      Contact( #iOTS_Frm_Prev_TTDown )
      Coil( #s130_StChkTTDwnRdyToRecv_T1 )
   END_RUNG
   RUNG wire#w1
      I_Contact( #s130_StChkTTDwnRdyToRecv_T1 )
      I_Contact( #iOTS_Frm_Prev_TTDown )
      Contact( #sTTDwn_90Pos_RX_Time )
      Coil( #s130_StChkTTDwnRdyToRecv_T2 )
   END_RUNG
   // the same network as SCL:
   #_w1 := #s130_StChkTTDwnRdyToRecv AND NOT #sStWtResetRel AND #sSst;
   #s130_StChkTTDwnRdyToRecv_T1 := #_w1 AND #iOTS_Frm_Prev_TTDown;
   #s130_StChkTTDwnRdyToRecv_T2 := #_w1 AND NOT #s130_StChkTTDwnRdyToRecv_T1 AND NOT #iOTS_Frm_Prev_TTDown AND #sTTDwn_90Pos_RX_Time;
END_REGION

REGION Network 49: STATE Num:130 StChkTTDwnRdyToRecv
   RUNG wire#powerrail
      Contact( #s130_StChkTTDwnRdyToRecv )
      wire#w1
      I_Contact( #sStWtResetRel )
      I_Contact( #s130_StChkTTDwnRdyToRecv_T1 )
      I_Contact( #s130_StChkTTDwnRdyToRecv_T2 )
      wire#w2
      Coil( #s130_StChkTTDwnRdyToRecv )
   END_RUNG
   RUNG wire#powerrail
      Contact( #s120_StWtForTTLck_T1 )
   END_RUNG wire#w1
   RUNG wire#w2
      { S7_GenerateENO := "TRUE" } Move(in := 130, out1 => #StateNo)
   END_RUNG
   // the same network as SCL:
   #s130_StChkTTDwnRdyToRecv := (#s130_StChkTTDwnRdyToRecv OR #s120_StWtForTTLck_T1) AND NOT #sStWtResetRel AND NOT #s130_StChkTTDwnRdyToRecv_T1 AND NOT #s130_StChkTTDwnRdyToRecv_T2;
   IF #s130_StChkTTDwnRdyToRecv THEN #StateNo := 130; END_IF;
END_REGION

REGION Network 50: Actions for STATE Num:130 StChkTTDwnRdyToRecv
   RUNG wire#powerrail
      Contact( #s130_StChkTTDwnRdyToRecv )
      Coil( #qRTR_Frm_TTDwn )
   END_RUNG
   // the same network as SCL:
   #qRTR_Frm_TTDwn := #s130_StChkTTDwnRdyToRecv;
END_REGION

REGION Network 51: Transition for STATE Num:140 StWtFrConveyorStrt
   RUNG wire#powerrail
      Contact( #s140_StWtFrConveyorStrt )
      I_Contact( #sStWtResetRel )
      Contact( #sSst )
      wire#w1
      Contact( #iPalletPrsnt_TTDown )
      Contact( #sPalletPrsntDebTTDown )
      Contact( #iRecvAreaClr_TTDown )
      wire#w2
      Coil( #s140_StWtFrConveyorStrt_T1 )
   END_RUNG
   RUNG wire#w1
      Contact( #sOTSFrmDwnTout )
   END_RUNG wire#w2
   // the same network as SCL:
   #s140_StWtFrConveyorStrt_T1 := #s140_StWtFrConveyorStrt AND NOT #sStWtResetRel AND #sSst AND ((#iPalletPrsnt_TTDown AND #sPalletPrsntDebTTDown AND #iRecvAreaClr_TTDown) OR #sOTSFrmDwnTout);
END_REGION

REGION Network 52: STATE Num:140 StWtFrConveyorStrt
   RUNG wire#powerrail
      Contact( #s140_StWtFrConveyorStrt )
      wire#w1
      I_Contact( #sStWtResetRel )
      I_Contact( #s140_StWtFrConveyorStrt_T1 )
      wire#w2
      Coil( #s140_StWtFrConveyorStrt )
   END_RUNG
   RUNG wire#powerrail
      Contact( #s130_StChkTTDwnRdyToRecv_T1 )
   END_RUNG wire#w1
   RUNG wire#powerrail
      Contact( #s130_StChkTTDwnRdyToRecv_T2 )
   END_RUNG wire#w1
   RUNG wire#w2
      { S7_GenerateENO := "TRUE" } Move(in := 140, out1 => #StateNo)
   END_RUNG
   // the same network as SCL:
   #s140_StWtFrConveyorStrt := (#s140_StWtFrConveyorStrt OR #s130_StChkTTDwnRdyToRecv_T1 OR #s130_StChkTTDwnRdyToRecv_T2) AND NOT #sStWtResetRel AND NOT #s140_StWtFrConveyorStrt_T1;
   IF #s140_StWtFrConveyorStrt THEN #StateNo := 140; END_IF;
END_REGION

REGION Network 53: Actions for STATE Num:140 StWtFrConveyorStrt
   RUNG wire#powerrail
      Contact( #s140_StWtFrConveyorStrt )
      Coil( #qConvRun_TTDown )
   END_RUNG
   // the same network as SCL:
   #qConvRun_TTDown := #s140_StWtFrConveyorStrt;
END_REGION

REGION Network 54: Transition for STATE Num:150 StChkNxtStRdyToRecvTTUp
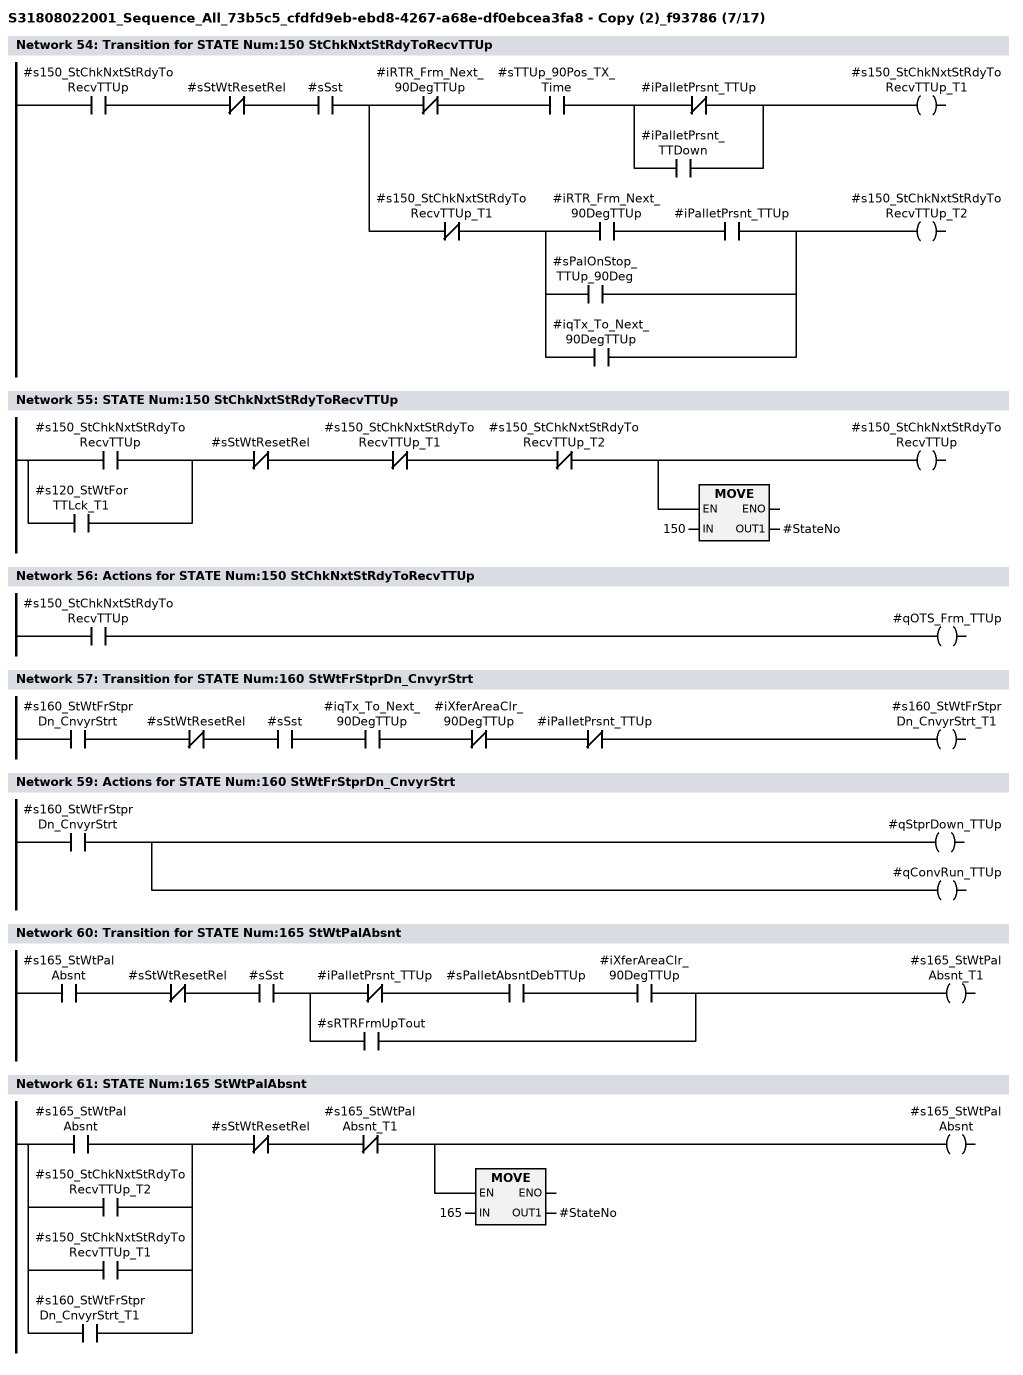
   RUNG wire#powerrail
      Contact( #s150_StChkNxtStRdyToRecvTTUp )
      I_Contact( #sStWtResetRel )
      Contact( #sSst )
      wire#w1
      I_Contact( #iRTR_Frm_Next_90DegTTUp )
      Contact( #sTTUp_90Pos_TX_Time )
      wire#w2
      I_Contact( #iPalletPrsnt_TTUp )
      wire#w3
      Coil( #s150_StChkNxtStRdyToRecvTTUp_T1 )
   END_RUNG
   RUNG wire#w2
      Contact( #iPalletPrsnt_TTDown )
   END_RUNG wire#w3
   RUNG wire#w1
      I_Contact( #s150_StChkNxtStRdyToRecvTTUp_T1 )
      wire#w4
      Contact( #iRTR_Frm_Next_90DegTTUp )
      Contact( #iPalletPrsnt_TTUp )
      wire#w5
      Coil( #s150_StChkNxtStRdyToRecvTTUp_T2 )
   END_RUNG
   RUNG wire#w4
      Contact( #sPalOnStop_TTUp_90Deg )
   END_RUNG wire#w5
   RUNG wire#w4
      Contact( #iqTx_To_Next_90DegTTUp )
   END_RUNG wire#w5
   // the same network as SCL:
   #_w1 := #s150_StChkNxtStRdyToRecvTTUp AND NOT #sStWtResetRel AND #sSst;
   #s150_StChkNxtStRdyToRecvTTUp_T1 := #_w1 AND NOT #iRTR_Frm_Next_90DegTTUp AND #sTTUp_90Pos_TX_Time AND (NOT #iPalletPrsnt_TTUp OR #iPalletPrsnt_TTDown);
   #s150_StChkNxtStRdyToRecvTTUp_T2 := #_w1 AND NOT #s150_StChkNxtStRdyToRecvTTUp_T1 AND ((#iRTR_Frm_Next_90DegTTUp AND #iPalletPrsnt_TTUp) OR #sPalOnStop_TTUp_90Deg OR #iqTx_To_Next_90DegTTUp);
END_REGION

REGION Network 55: STATE Num:150 StChkNxtStRdyToRecvTTUp
   RUNG wire#powerrail
      Contact( #s150_StChkNxtStRdyToRecvTTUp )
      wire#w1
      I_Contact( #sStWtResetRel )
      I_Contact( #s150_StChkNxtStRdyToRecvTTUp_T1 )
      I_Contact( #s150_StChkNxtStRdyToRecvTTUp_T2 )
      wire#w2
      Coil( #s150_StChkNxtStRdyToRecvTTUp )
   END_RUNG
   RUNG wire#powerrail
      Contact( #s120_StWtForTTLck_T1 )
   END_RUNG wire#w1
   RUNG wire#w2
      { S7_GenerateENO := "TRUE" } Move(in := 150, out1 => #StateNo)
   END_RUNG
   // the same network as SCL:
   #s150_StChkNxtStRdyToRecvTTUp := (#s150_StChkNxtStRdyToRecvTTUp OR #s120_StWtForTTLck_T1) AND NOT #sStWtResetRel AND NOT #s150_StChkNxtStRdyToRecvTTUp_T1 AND NOT #s150_StChkNxtStRdyToRecvTTUp_T2;
   IF #s150_StChkNxtStRdyToRecvTTUp THEN #StateNo := 150; END_IF;
END_REGION

REGION Network 56: Actions for STATE Num:150 StChkNxtStRdyToRecvTTUp
   RUNG wire#powerrail
      Contact( #s150_StChkNxtStRdyToRecvTTUp )
      Coil( #qOTS_Frm_TTUp )
   END_RUNG
   // the same network as SCL:
   #qOTS_Frm_TTUp := #s150_StChkNxtStRdyToRecvTTUp;
END_REGION

REGION Network 57: Transition for STATE Num:160 StWtFrStprDn_CnvyrStrt
   RUNG wire#powerrail
      Contact( #s160_StWtFrStprDn_CnvyrStrt )
      I_Contact( #sStWtResetRel )
      Contact( #sSst )
      Contact( #iqTx_To_Next_90DegTTUp )
      I_Contact( #iXferAreaClr_90DegTTUp )
      I_Contact( #iPalletPrsnt_TTUp )
      Coil( #s160_StWtFrStprDn_CnvyrStrt_T1 )
   END_RUNG
   // the same network as SCL:
   #s160_StWtFrStprDn_CnvyrStrt_T1 := #s160_StWtFrStprDn_CnvyrStrt AND NOT #sStWtResetRel AND #sSst AND #iqTx_To_Next_90DegTTUp AND NOT #iXferAreaClr_90DegTTUp AND NOT #iPalletPrsnt_TTUp;
END_REGION

NETWORK
TITLE = STATE Num:160 StWtFrStprDn_CnvyrStrt
      A(;
      O     #s160_StWtFrStprDn_CnvyrStrt;
//wrong transition variable removed
      );
      AN    #sStWtResetRel;
      AN    #s160_StWtFrStprDn_CnvyrStrt_T1;
      =     %L1.0;
      A     %L1.0;
      BLD   102;
      =     #s160_StWtFrStprDn_CnvyrStrt;
      A     %L1.0;
      JNB   Label_19;
      L     160;
      T     #StateNo;
Label_19:NOP   0;

REGION Network 59: Actions for STATE Num:160 StWtFrStprDn_CnvyrStrt
   RUNG wire#powerrail
      Contact( #s160_StWtFrStprDn_CnvyrStrt )
      wire#w1
      Coil( #qStprDown_TTUp )
   END_RUNG
   RUNG wire#w1
      Coil( #qConvRun_TTUp )
   END_RUNG
   // the same network as SCL:
   #qStprDown_TTUp := #s160_StWtFrStprDn_CnvyrStrt;
   #qConvRun_TTUp := #s160_StWtFrStprDn_CnvyrStrt;
END_REGION

REGION Network 60: Transition for STATE Num:165 StWtPalAbsnt
   RUNG wire#powerrail
      Contact( #s165_StWtPalAbsnt )
      I_Contact( #sStWtResetRel )
      Contact( #sSst )
      wire#w1
      I_Contact( #iPalletPrsnt_TTUp )
      Contact( #sPalletAbsntDebTTUp )
      Contact( #iXferAreaClr_90DegTTUp )
      wire#w2
      Coil( #s165_StWtPalAbsnt_T1 )
   END_RUNG
   RUNG wire#w1
      Contact( #sRTRFrmUpTout )
   END_RUNG wire#w2
   // the same network as SCL:
   #s165_StWtPalAbsnt_T1 := #s165_StWtPalAbsnt AND NOT #sStWtResetRel AND #sSst AND ((NOT #iPalletPrsnt_TTUp AND #sPalletAbsntDebTTUp AND #iXferAreaClr_90DegTTUp) OR #sRTRFrmUpTout);
END_REGION

REGION Network 61: STATE Num:165 StWtPalAbsnt
   RUNG wire#powerrail
      Contact( #s165_StWtPalAbsnt )
      wire#w1
      I_Contact( #sStWtResetRel )
      I_Contact( #s165_StWtPalAbsnt_T1 )
      wire#w2
      Coil( #s165_StWtPalAbsnt )
   END_RUNG
   RUNG wire#powerrail
      Contact( #s150_StChkNxtStRdyToRecvTTUp_T2 )
   END_RUNG wire#w1
   RUNG wire#powerrail
      Contact( #s150_StChkNxtStRdyToRecvTTUp_T1 )
   END_RUNG wire#w1
   RUNG wire#powerrail
      Contact( #s160_StWtFrStprDn_CnvyrStrt_T1 )
   END_RUNG wire#w1
   RUNG wire#w2
      { S7_GenerateENO := "TRUE" } Move(in := 165, out1 => #StateNo)
   END_RUNG
   // the same network as SCL:
   #s165_StWtPalAbsnt := (#s165_StWtPalAbsnt OR #s150_StChkNxtStRdyToRecvTTUp_T2 OR #s150_StChkNxtStRdyToRecvTTUp_T1 OR #s160_StWtFrStprDn_CnvyrStrt_T1) AND NOT #sStWtResetRel AND NOT #s165_StWtPalAbsnt_T1;
   IF #s165_StWtPalAbsnt THEN #StateNo := 165; END_IF;
END_REGION

REGION Network 62: Actions for STATE Num:165 StWtPalAbsnt
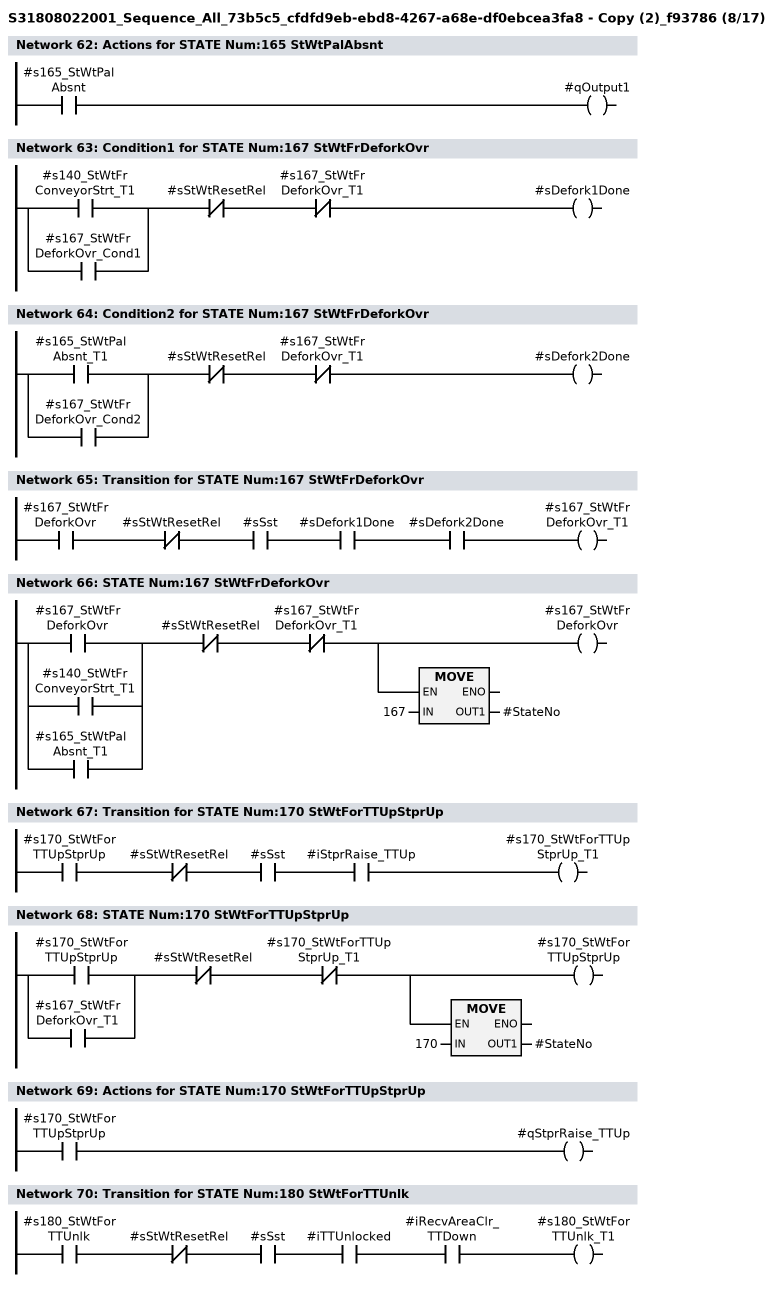
   RUNG wire#powerrail
      Contact( #s165_StWtPalAbsnt )
      Coil( #qOutput1 )
   END_RUNG
   // the same network as SCL:
   #qOutput1 := #s165_StWtPalAbsnt;
END_REGION

REGION Network 63: Condition1 for STATE Num:167 StWtFrDeforkOvr
   RUNG wire#powerrail
      Contact( #s140_StWtFrConveyorStrt_T1 )
      wire#w1
      I_Contact( #sStWtResetRel )
      I_Contact( #s167_StWtFrDeforkOvr_T1 )
      Coil( #sDefork1Done )
   END_RUNG
   RUNG wire#powerrail
      Contact( #s167_StWtFrDeforkOvr_Cond1 )
   END_RUNG wire#w1
   // the same network as SCL:
   #sDefork1Done := (#s140_StWtFrConveyorStrt_T1 OR #s167_StWtFrDeforkOvr_Cond1) AND NOT #sStWtResetRel AND NOT #s167_StWtFrDeforkOvr_T1;
END_REGION

REGION Network 64: Condition2 for STATE Num:167 StWtFrDeforkOvr
   RUNG wire#powerrail
      Contact( #s165_StWtPalAbsnt_T1 )
      wire#w1
      I_Contact( #sStWtResetRel )
      I_Contact( #s167_StWtFrDeforkOvr_T1 )
      Coil( #sDefork2Done )
   END_RUNG
   RUNG wire#powerrail
      Contact( #s167_StWtFrDeforkOvr_Cond2 )
   END_RUNG wire#w1
   // the same network as SCL:
   #sDefork2Done := (#s165_StWtPalAbsnt_T1 OR #s167_StWtFrDeforkOvr_Cond2) AND NOT #sStWtResetRel AND NOT #s167_StWtFrDeforkOvr_T1;
END_REGION

REGION Network 65: Transition for STATE Num:167 StWtFrDeforkOvr
   RUNG wire#powerrail
      Contact( #s167_StWtFrDeforkOvr )
      I_Contact( #sStWtResetRel )
      Contact( #sSst )
      Contact( #sDefork1Done )
      Contact( #sDefork2Done )
      Coil( #s167_StWtFrDeforkOvr_T1 )
   END_RUNG
   // the same network as SCL:
   #s167_StWtFrDeforkOvr_T1 := #s167_StWtFrDeforkOvr AND NOT #sStWtResetRel AND #sSst AND #sDefork1Done AND #sDefork2Done;
END_REGION

REGION Network 66: STATE Num:167 StWtFrDeforkOvr
   RUNG wire#powerrail
      Contact( #s167_StWtFrDeforkOvr )
      wire#w1
      I_Contact( #sStWtResetRel )
      I_Contact( #s167_StWtFrDeforkOvr_T1 )
      wire#w2
      Coil( #s167_StWtFrDeforkOvr )
   END_RUNG
   RUNG wire#powerrail
      Contact( #s140_StWtFrConveyorStrt_T1 )
   END_RUNG wire#w1
   RUNG wire#powerrail
      Contact( #s165_StWtPalAbsnt_T1 )
   END_RUNG wire#w1
   RUNG wire#w2
      { S7_GenerateENO := "TRUE" } Move(in := 167, out1 => #StateNo)
   END_RUNG
   // the same network as SCL:
   #s167_StWtFrDeforkOvr := (#s167_StWtFrDeforkOvr OR #s140_StWtFrConveyorStrt_T1 OR #s165_StWtPalAbsnt_T1) AND NOT #sStWtResetRel AND NOT #s167_StWtFrDeforkOvr_T1;
   IF #s167_StWtFrDeforkOvr THEN #StateNo := 167; END_IF;
END_REGION

REGION Network 67: Transition for STATE Num:170 StWtForTTUpStprUp
   RUNG wire#powerrail
      Contact( #s170_StWtForTTUpStprUp )
      I_Contact( #sStWtResetRel )
      Contact( #sSst )
      Contact( #iStprRaise_TTUp )
      Coil( #s170_StWtForTTUpStprUp_T1 )
   END_RUNG
   // the same network as SCL:
   #s170_StWtForTTUpStprUp_T1 := #s170_StWtForTTUpStprUp AND NOT #sStWtResetRel AND #sSst AND #iStprRaise_TTUp;
END_REGION

REGION Network 68: STATE Num:170 StWtForTTUpStprUp
   RUNG wire#powerrail
      Contact( #s170_StWtForTTUpStprUp )
      wire#w1
      I_Contact( #sStWtResetRel )
      I_Contact( #s170_StWtForTTUpStprUp_T1 )
      wire#w2
      Coil( #s170_StWtForTTUpStprUp )
   END_RUNG
   RUNG wire#powerrail
      Contact( #s167_StWtFrDeforkOvr_T1 )
   END_RUNG wire#w1
   RUNG wire#w2
      { S7_GenerateENO := "TRUE" } Move(in := 170, out1 => #StateNo)
   END_RUNG
   // the same network as SCL:
   #s170_StWtForTTUpStprUp := (#s170_StWtForTTUpStprUp OR #s167_StWtFrDeforkOvr_T1) AND NOT #sStWtResetRel AND NOT #s170_StWtForTTUpStprUp_T1;
   IF #s170_StWtForTTUpStprUp THEN #StateNo := 170; END_IF;
END_REGION

REGION Network 69: Actions for STATE Num:170 StWtForTTUpStprUp
   RUNG wire#powerrail
      Contact( #s170_StWtForTTUpStprUp )
      Coil( #qStprRaise_TTUp )
   END_RUNG
   // the same network as SCL:
   #qStprRaise_TTUp := #s170_StWtForTTUpStprUp;
END_REGION

REGION Network 70: Transition for STATE Num:180 StWtForTTUnlk
   RUNG wire#powerrail
      Contact( #s180_StWtForTTUnlk )
      I_Contact( #sStWtResetRel )
      Contact( #sSst )
      Contact( #iTTUnlocked )
      Contact( #iRecvAreaClr_TTDown )
      Coil( #s180_StWtForTTUnlk_T1 )
   END_RUNG
   // the same network as SCL:
   #s180_StWtForTTUnlk_T1 := #s180_StWtForTTUnlk AND NOT #sStWtResetRel AND #sSst AND #iTTUnlocked AND #iRecvAreaClr_TTDown;
END_REGION

REGION Network 71: STATE Num:180 StWtForTTUnlk
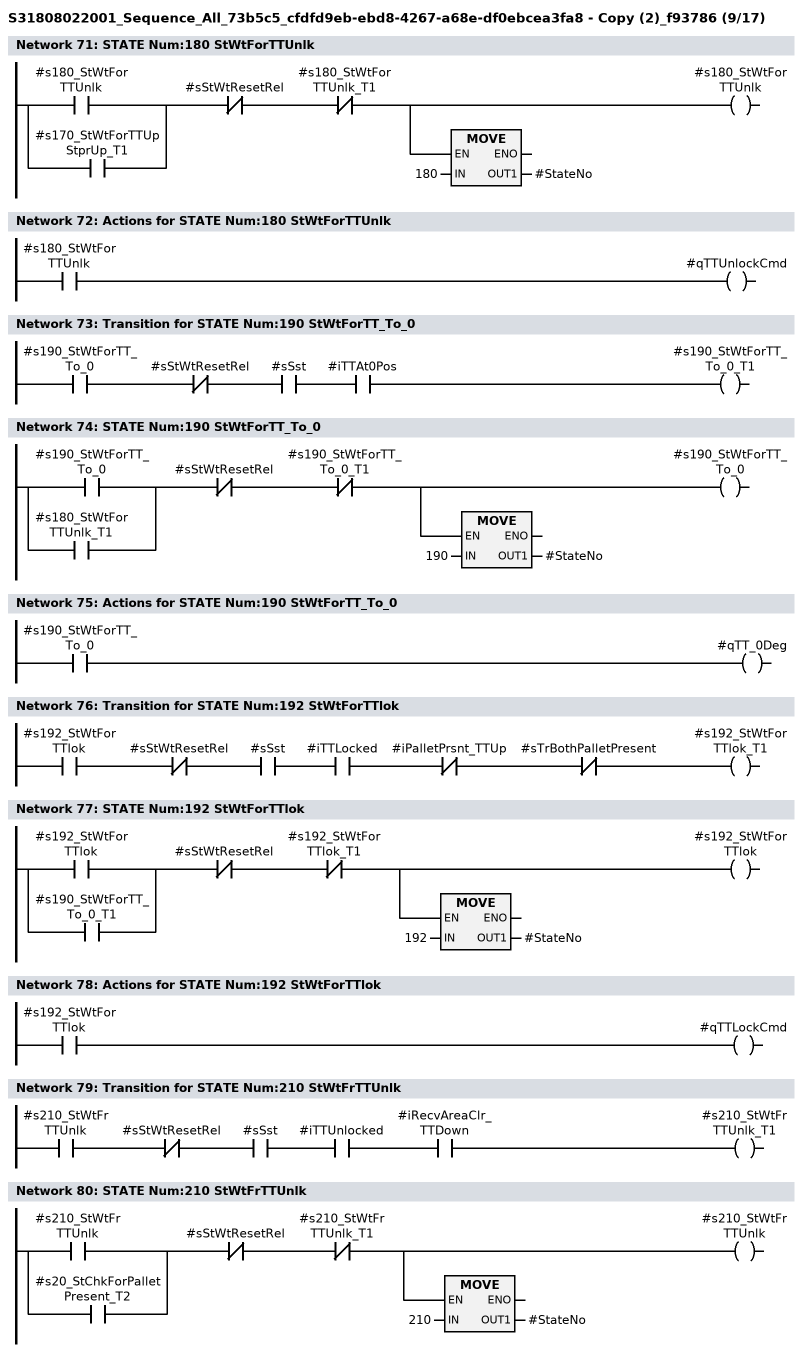
   RUNG wire#powerrail
      Contact( #s180_StWtForTTUnlk )
      wire#w1
      I_Contact( #sStWtResetRel )
      I_Contact( #s180_StWtForTTUnlk_T1 )
      wire#w2
      Coil( #s180_StWtForTTUnlk )
   END_RUNG
   RUNG wire#powerrail
      Contact( #s170_StWtForTTUpStprUp_T1 )
   END_RUNG wire#w1
   RUNG wire#w2
      { S7_GenerateENO := "TRUE" } Move(in := 180, out1 => #StateNo)
   END_RUNG
   // the same network as SCL:
   #s180_StWtForTTUnlk := (#s180_StWtForTTUnlk OR #s170_StWtForTTUpStprUp_T1) AND NOT #sStWtResetRel AND NOT #s180_StWtForTTUnlk_T1;
   IF #s180_StWtForTTUnlk THEN #StateNo := 180; END_IF;
END_REGION

REGION Network 72: Actions for STATE Num:180 StWtForTTUnlk
   RUNG wire#powerrail
      Contact( #s180_StWtForTTUnlk )
      Coil( #qTTUnlockCmd )
   END_RUNG
   // the same network as SCL:
   #qTTUnlockCmd := #s180_StWtForTTUnlk;
END_REGION

REGION Network 73: Transition for STATE Num:190 StWtForTT_To_0
   RUNG wire#powerrail
      Contact( #s190_StWtForTT_To_0 )
      I_Contact( #sStWtResetRel )
      Contact( #sSst )
      Contact( #iTTAt0Pos )
      Coil( #s190_StWtForTT_To_0_T1 )
   END_RUNG
   // the same network as SCL:
   #s190_StWtForTT_To_0_T1 := #s190_StWtForTT_To_0 AND NOT #sStWtResetRel AND #sSst AND #iTTAt0Pos;
END_REGION

REGION Network 74: STATE Num:190 StWtForTT_To_0
   RUNG wire#powerrail
      Contact( #s190_StWtForTT_To_0 )
      wire#w1
      I_Contact( #sStWtResetRel )
      I_Contact( #s190_StWtForTT_To_0_T1 )
      wire#w2
      Coil( #s190_StWtForTT_To_0 )
   END_RUNG
   RUNG wire#powerrail
      Contact( #s180_StWtForTTUnlk_T1 )
   END_RUNG wire#w1
   RUNG wire#w2
      { S7_GenerateENO := "TRUE" } Move(in := 190, out1 => #StateNo)
   END_RUNG
   // the same network as SCL:
   #s190_StWtForTT_To_0 := (#s190_StWtForTT_To_0 OR #s180_StWtForTTUnlk_T1) AND NOT #sStWtResetRel AND NOT #s190_StWtForTT_To_0_T1;
   IF #s190_StWtForTT_To_0 THEN #StateNo := 190; END_IF;
END_REGION

REGION Network 75: Actions for STATE Num:190 StWtForTT_To_0
   RUNG wire#powerrail
      Contact( #s190_StWtForTT_To_0 )
      Coil( #qTT_0Deg )
   END_RUNG
   // the same network as SCL:
   #qTT_0Deg := #s190_StWtForTT_To_0;
END_REGION

REGION Network 76: Transition for STATE Num:192 StWtForTTlok
   RUNG wire#powerrail
      Contact( #s192_StWtForTTlok )
      I_Contact( #sStWtResetRel )
      Contact( #sSst )
      Contact( #iTTLocked )
      I_Contact( #iPalletPrsnt_TTUp )
      I_Contact( #sTrBothPalletPresent )
      Coil( #s192_StWtForTTlok_T1 )
   END_RUNG
   // the same network as SCL:
   #s192_StWtForTTlok_T1 := #s192_StWtForTTlok AND NOT #sStWtResetRel AND #sSst AND #iTTLocked AND NOT #iPalletPrsnt_TTUp AND NOT #sTrBothPalletPresent;
END_REGION

REGION Network 77: STATE Num:192 StWtForTTlok
   RUNG wire#powerrail
      Contact( #s192_StWtForTTlok )
      wire#w1
      I_Contact( #sStWtResetRel )
      I_Contact( #s192_StWtForTTlok_T1 )
      wire#w2
      Coil( #s192_StWtForTTlok )
   END_RUNG
   RUNG wire#powerrail
      Contact( #s190_StWtForTT_To_0_T1 )
   END_RUNG wire#w1
   RUNG wire#w2
      { S7_GenerateENO := "TRUE" } Move(in := 192, out1 => #StateNo)
   END_RUNG
   // the same network as SCL:
   #s192_StWtForTTlok := (#s192_StWtForTTlok OR #s190_StWtForTT_To_0_T1) AND NOT #sStWtResetRel AND NOT #s192_StWtForTTlok_T1;
   IF #s192_StWtForTTlok THEN #StateNo := 192; END_IF;
END_REGION

REGION Network 78: Actions for STATE Num:192 StWtForTTlok
   RUNG wire#powerrail
      Contact( #s192_StWtForTTlok )
      Coil( #qTTLockCmd )
   END_RUNG
   // the same network as SCL:
   #qTTLockCmd := #s192_StWtForTTlok;
END_REGION

REGION Network 79: Transition for STATE Num:210 StWtFrTTUnlk
   RUNG wire#powerrail
      Contact( #s210_StWtFrTTUnlk )
      I_Contact( #sStWtResetRel )
      Contact( #sSst )
      Contact( #iTTUnlocked )
      Contact( #iRecvAreaClr_TTDown )
      Coil( #s210_StWtFrTTUnlk_T1 )
   END_RUNG
   // the same network as SCL:
   #s210_StWtFrTTUnlk_T1 := #s210_StWtFrTTUnlk AND NOT #sStWtResetRel AND #sSst AND #iTTUnlocked AND #iRecvAreaClr_TTDown;
END_REGION

REGION Network 80: STATE Num:210 StWtFrTTUnlk
   RUNG wire#powerrail
      Contact( #s210_StWtFrTTUnlk )
      wire#w1
      I_Contact( #sStWtResetRel )
      I_Contact( #s210_StWtFrTTUnlk_T1 )
      wire#w2
      Coil( #s210_StWtFrTTUnlk )
   END_RUNG
   RUNG wire#powerrail
      Contact( #s20_StChkForPalletPresent_T2 )
   END_RUNG wire#w1
   RUNG wire#w2
      { S7_GenerateENO := "TRUE" } Move(in := 210, out1 => #StateNo)
   END_RUNG
   // the same network as SCL:
   #s210_StWtFrTTUnlk := (#s210_StWtFrTTUnlk OR #s20_StChkForPalletPresent_T2) AND NOT #sStWtResetRel AND NOT #s210_StWtFrTTUnlk_T1;
   IF #s210_StWtFrTTUnlk THEN #StateNo := 210; END_IF;
END_REGION

REGION Network 81: Actions for STATE Num:210 StWtFrTTUnlk
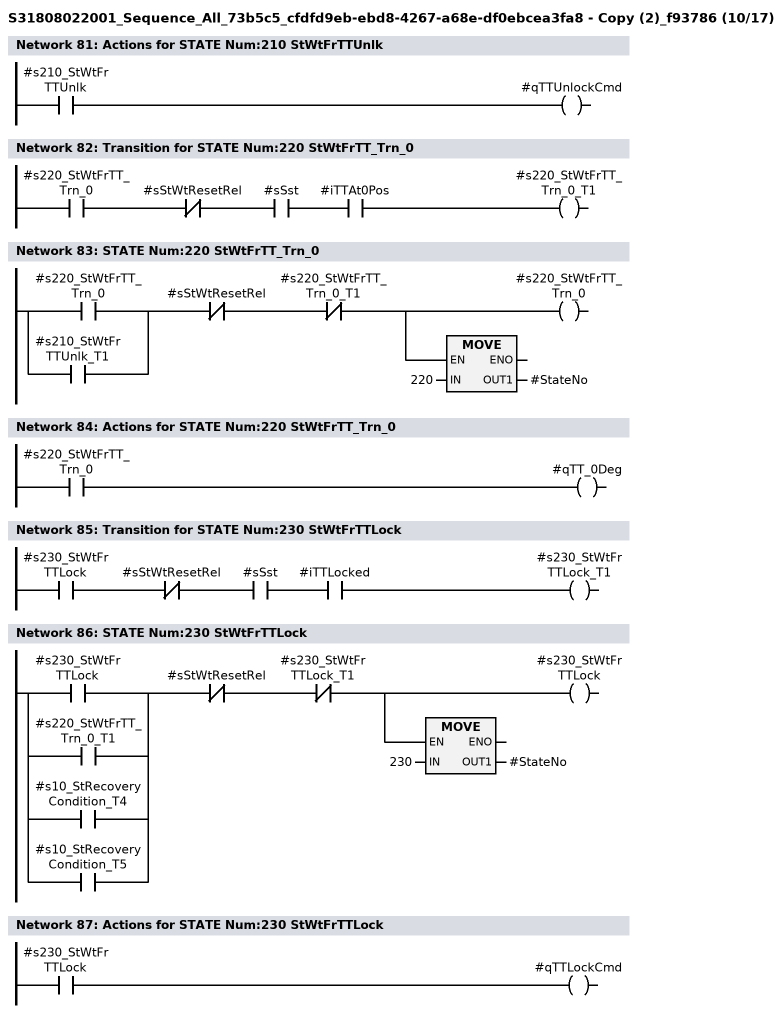
   RUNG wire#powerrail
      Contact( #s210_StWtFrTTUnlk )
      Coil( #qTTUnlockCmd )
   END_RUNG
   // the same network as SCL:
   #qTTUnlockCmd := #s210_StWtFrTTUnlk;
END_REGION

REGION Network 82: Transition for STATE Num:220 StWtFrTT_Trn_0
   RUNG wire#powerrail
      Contact( #s220_StWtFrTT_Trn_0 )
      I_Contact( #sStWtResetRel )
      Contact( #sSst )
      Contact( #iTTAt0Pos )
      Coil( #s220_StWtFrTT_Trn_0_T1 )
   END_RUNG
   // the same network as SCL:
   #s220_StWtFrTT_Trn_0_T1 := #s220_StWtFrTT_Trn_0 AND NOT #sStWtResetRel AND #sSst AND #iTTAt0Pos;
END_REGION

REGION Network 83: STATE Num:220 StWtFrTT_Trn_0
   RUNG wire#powerrail
      Contact( #s220_StWtFrTT_Trn_0 )
      wire#w1
      I_Contact( #sStWtResetRel )
      I_Contact( #s220_StWtFrTT_Trn_0_T1 )
      wire#w2
      Coil( #s220_StWtFrTT_Trn_0 )
   END_RUNG
   RUNG wire#powerrail
      Contact( #s210_StWtFrTTUnlk_T1 )
   END_RUNG wire#w1
   RUNG wire#w2
      { S7_GenerateENO := "TRUE" } Move(in := 220, out1 => #StateNo)
   END_RUNG
   // the same network as SCL:
   #s220_StWtFrTT_Trn_0 := (#s220_StWtFrTT_Trn_0 OR #s210_StWtFrTTUnlk_T1) AND NOT #sStWtResetRel AND NOT #s220_StWtFrTT_Trn_0_T1;
   IF #s220_StWtFrTT_Trn_0 THEN #StateNo := 220; END_IF;
END_REGION

REGION Network 84: Actions for STATE Num:220 StWtFrTT_Trn_0
   RUNG wire#powerrail
      Contact( #s220_StWtFrTT_Trn_0 )
      Coil( #qTT_0Deg )
   END_RUNG
   // the same network as SCL:
   #qTT_0Deg := #s220_StWtFrTT_Trn_0;
END_REGION

REGION Network 85: Transition for STATE Num:230 StWtFrTTLock
   RUNG wire#powerrail
      Contact( #s230_StWtFrTTLock )
      I_Contact( #sStWtResetRel )
      Contact( #sSst )
      Contact( #iTTLocked )
      Coil( #s230_StWtFrTTLock_T1 )
   END_RUNG
   // the same network as SCL:
   #s230_StWtFrTTLock_T1 := #s230_StWtFrTTLock AND NOT #sStWtResetRel AND #sSst AND #iTTLocked;
END_REGION

REGION Network 86: STATE Num:230 StWtFrTTLock
   RUNG wire#powerrail
      Contact( #s230_StWtFrTTLock )
      wire#w1
      I_Contact( #sStWtResetRel )
      I_Contact( #s230_StWtFrTTLock_T1 )
      wire#w2
      Coil( #s230_StWtFrTTLock )
   END_RUNG
   RUNG wire#powerrail
      Contact( #s220_StWtFrTT_Trn_0_T1 )
   END_RUNG wire#w1
   RUNG wire#powerrail
      Contact( #s10_StRecoveryCondition_T4 )
   END_RUNG wire#w1
   RUNG wire#powerrail
      Contact( #s10_StRecoveryCondition_T5 )
   END_RUNG wire#w1
   RUNG wire#w2
      { S7_GenerateENO := "TRUE" } Move(in := 230, out1 => #StateNo)
   END_RUNG
   // the same network as SCL:
   #s230_StWtFrTTLock := (#s230_StWtFrTTLock OR #s220_StWtFrTT_Trn_0_T1 OR #s10_StRecoveryCondition_T4 OR #s10_StRecoveryCondition_T5) AND NOT #sStWtResetRel AND NOT #s230_StWtFrTTLock_T1;
   IF #s230_StWtFrTTLock THEN #StateNo := 230; END_IF;
END_REGION

REGION Network 87: Actions for STATE Num:230 StWtFrTTLock
   RUNG wire#powerrail
      Contact( #s230_StWtFrTTLock )
      Coil( #qTTLockCmd )
   END_RUNG
   // the same network as SCL:
   #qTTLockCmd := #s230_StWtFrTTLock;
END_REGION

REGION Network 88: Transition for STATE Num:240 StWtFRTRNxtStnTTDown
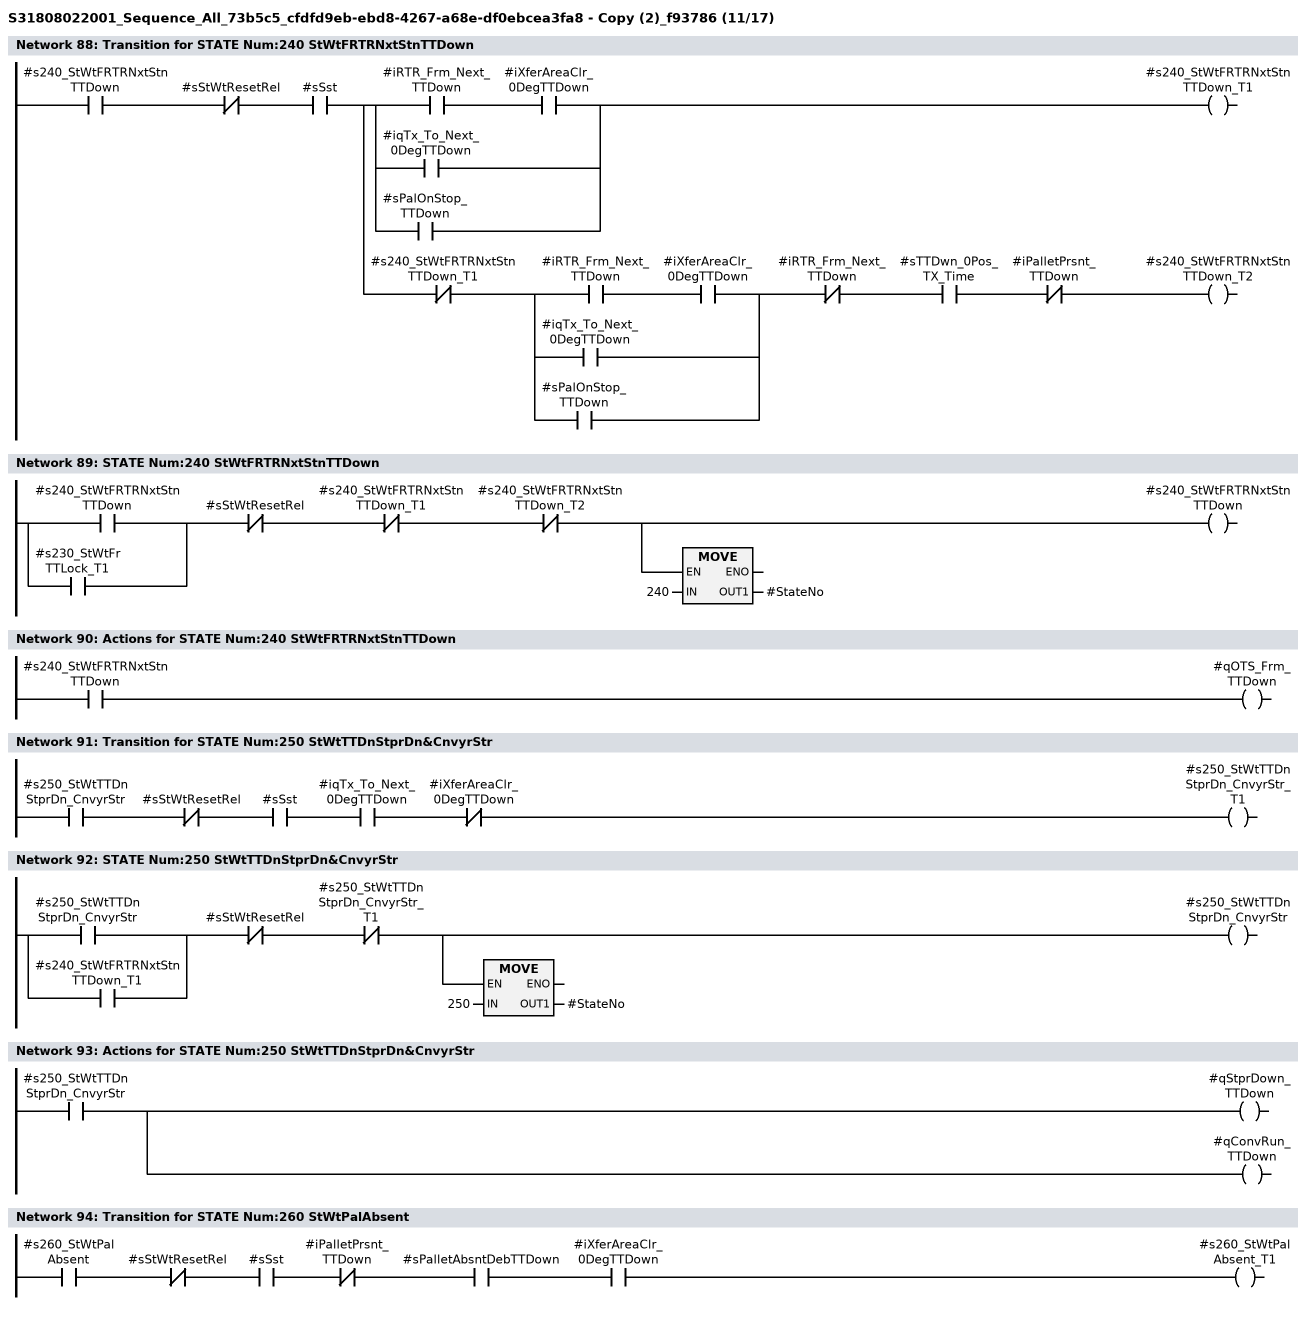
   RUNG wire#powerrail
      Contact( #s240_StWtFRTRNxtStnTTDown )
      I_Contact( #sStWtResetRel )
      Contact( #sSst )
      wire#w1
      Contact( #iRTR_Frm_Next_TTDown )
      Contact( #iXferAreaClr_0DegTTDown )
      wire#w2
      Coil( #s240_StWtFRTRNxtStnTTDown_T1 )
   END_RUNG
   RUNG wire#w1
      Contact( #iqTx_To_Next_0DegTTDown )
   END_RUNG wire#w2
   RUNG wire#w1
      Contact( #sPalOnStop_TTDown )
   END_RUNG wire#w2
   RUNG wire#w1
      I_Contact( #s240_StWtFRTRNxtStnTTDown_T1 )
      wire#w3
      Contact( #iRTR_Frm_Next_TTDown )
      Contact( #iXferAreaClr_0DegTTDown )
      wire#w4
      I_Contact( #iRTR_Frm_Next_TTDown )
      Contact( #sTTDwn_0Pos_TX_Time )
      I_Contact( #iPalletPrsnt_TTDown )
      Coil( #s240_StWtFRTRNxtStnTTDown_T2 )
   END_RUNG
   RUNG wire#w3
      Contact( #iqTx_To_Next_0DegTTDown )
   END_RUNG wire#w4
   RUNG wire#w3
      Contact( #sPalOnStop_TTDown )
   END_RUNG wire#w4
   // the same network as SCL:
   #_w1 := #s240_StWtFRTRNxtStnTTDown AND NOT #sStWtResetRel AND #sSst;
   #s240_StWtFRTRNxtStnTTDown_T1 := #_w1 AND ((#iRTR_Frm_Next_TTDown AND #iXferAreaClr_0DegTTDown) OR #iqTx_To_Next_0DegTTDown OR #sPalOnStop_TTDown);
   #s240_StWtFRTRNxtStnTTDown_T2 := #_w1 AND NOT #s240_StWtFRTRNxtStnTTDown_T1 AND ((#iRTR_Frm_Next_TTDown AND #iXferAreaClr_0DegTTDown) OR #iqTx_To_Next_0DegTTDown OR #sPalOnStop_TTDown) AND NOT #iRTR_Frm_Next_TTDown AND #sTTDwn_0Pos_TX_Time AND NOT #iPalletPrsnt_TTDown;
END_REGION

REGION Network 89: STATE Num:240 StWtFRTRNxtStnTTDown
   RUNG wire#powerrail
      Contact( #s240_StWtFRTRNxtStnTTDown )
      wire#w1
      I_Contact( #sStWtResetRel )
      I_Contact( #s240_StWtFRTRNxtStnTTDown_T1 )
      I_Contact( #s240_StWtFRTRNxtStnTTDown_T2 )
      wire#w2
      Coil( #s240_StWtFRTRNxtStnTTDown )
   END_RUNG
   RUNG wire#powerrail
      Contact( #s230_StWtFrTTLock_T1 )
   END_RUNG wire#w1
   RUNG wire#w2
      { S7_GenerateENO := "TRUE" } Move(in := 240, out1 => #StateNo)
   END_RUNG
   // the same network as SCL:
   #s240_StWtFRTRNxtStnTTDown := (#s240_StWtFRTRNxtStnTTDown OR #s230_StWtFrTTLock_T1) AND NOT #sStWtResetRel AND NOT #s240_StWtFRTRNxtStnTTDown_T1 AND NOT #s240_StWtFRTRNxtStnTTDown_T2;
   IF #s240_StWtFRTRNxtStnTTDown THEN #StateNo := 240; END_IF;
END_REGION

REGION Network 90: Actions for STATE Num:240 StWtFRTRNxtStnTTDown
   RUNG wire#powerrail
      Contact( #s240_StWtFRTRNxtStnTTDown )
      Coil( #qOTS_Frm_TTDown )
   END_RUNG
   // the same network as SCL:
   #qOTS_Frm_TTDown := #s240_StWtFRTRNxtStnTTDown;
END_REGION

REGION Network 91: Transition for STATE Num:250 StWtTTDnStprDn&CnvyrStr
   RUNG wire#powerrail
      Contact( #s250_StWtTTDnStprDn_CnvyrStr )
      I_Contact( #sStWtResetRel )
      Contact( #sSst )
      Contact( #iqTx_To_Next_0DegTTDown )
      I_Contact( #iXferAreaClr_0DegTTDown )
      Coil( #s250_StWtTTDnStprDn_CnvyrStr_T1 )
   END_RUNG
   // the same network as SCL:
   #s250_StWtTTDnStprDn_CnvyrStr_T1 := #s250_StWtTTDnStprDn_CnvyrStr AND NOT #sStWtResetRel AND #sSst AND #iqTx_To_Next_0DegTTDown AND NOT #iXferAreaClr_0DegTTDown;
END_REGION

REGION Network 92: STATE Num:250 StWtTTDnStprDn&CnvyrStr
   RUNG wire#powerrail
      Contact( #s250_StWtTTDnStprDn_CnvyrStr )
      wire#w1
      I_Contact( #sStWtResetRel )
      I_Contact( #s250_StWtTTDnStprDn_CnvyrStr_T1 )
      wire#w2
      Coil( #s250_StWtTTDnStprDn_CnvyrStr )
   END_RUNG
   RUNG wire#powerrail
      Contact( #s240_StWtFRTRNxtStnTTDown_T1 )
   END_RUNG wire#w1
   RUNG wire#w2
      { S7_GenerateENO := "TRUE" } Move(in := 250, out1 => #StateNo)
   END_RUNG
   // the same network as SCL:
   #s250_StWtTTDnStprDn_CnvyrStr := (#s250_StWtTTDnStprDn_CnvyrStr OR #s240_StWtFRTRNxtStnTTDown_T1) AND NOT #sStWtResetRel AND NOT #s250_StWtTTDnStprDn_CnvyrStr_T1;
   IF #s250_StWtTTDnStprDn_CnvyrStr THEN #StateNo := 250; END_IF;
END_REGION

REGION Network 93: Actions for STATE Num:250 StWtTTDnStprDn&CnvyrStr
   RUNG wire#powerrail
      Contact( #s250_StWtTTDnStprDn_CnvyrStr )
      wire#w1
      Coil( #qStprDown_TTDown )
   END_RUNG
   RUNG wire#w1
      Coil( #qConvRun_TTDown )
   END_RUNG
   // the same network as SCL:
   #qStprDown_TTDown := #s250_StWtTTDnStprDn_CnvyrStr;
   #qConvRun_TTDown := #s250_StWtTTDnStprDn_CnvyrStr;
END_REGION

REGION Network 94: Transition for STATE Num:260 StWtPalAbsent
   RUNG wire#powerrail
      Contact( #s260_StWtPalAbsent )
      I_Contact( #sStWtResetRel )
      Contact( #sSst )
      I_Contact( #iPalletPrsnt_TTDown )
      Contact( #sPalletAbsntDebTTDown )
      Contact( #iXferAreaClr_0DegTTDown )
      Coil( #s260_StWtPalAbsent_T1 )
   END_RUNG
   // the same network as SCL:
   #s260_StWtPalAbsent_T1 := #s260_StWtPalAbsent AND NOT #sStWtResetRel AND #sSst AND NOT #iPalletPrsnt_TTDown AND #sPalletAbsntDebTTDown AND #iXferAreaClr_0DegTTDown;
END_REGION

REGION Network 95: STATE Num:260 StWtPalAbsent
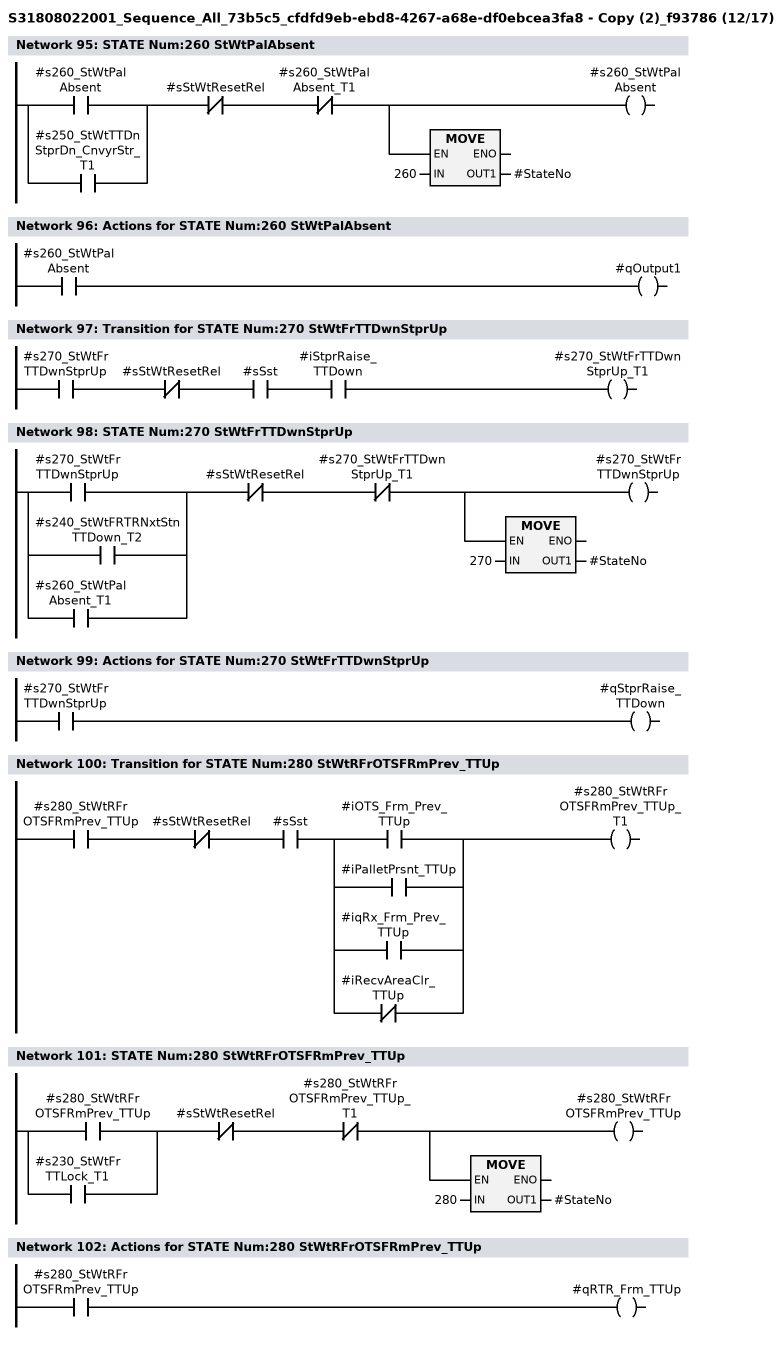
   RUNG wire#powerrail
      Contact( #s260_StWtPalAbsent )
      wire#w1
      I_Contact( #sStWtResetRel )
      I_Contact( #s260_StWtPalAbsent_T1 )
      wire#w2
      Coil( #s260_StWtPalAbsent )
   END_RUNG
   RUNG wire#powerrail
      Contact( #s250_StWtTTDnStprDn_CnvyrStr_T1 )
   END_RUNG wire#w1
   RUNG wire#w2
      { S7_GenerateENO := "TRUE" } Move(in := 260, out1 => #StateNo)
   END_RUNG
   // the same network as SCL:
   #s260_StWtPalAbsent := (#s260_StWtPalAbsent OR #s250_StWtTTDnStprDn_CnvyrStr_T1) AND NOT #sStWtResetRel AND NOT #s260_StWtPalAbsent_T1;
   IF #s260_StWtPalAbsent THEN #StateNo := 260; END_IF;
END_REGION

REGION Network 96: Actions for STATE Num:260 StWtPalAbsent
   RUNG wire#powerrail
      Contact( #s260_StWtPalAbsent )
      Coil( #qOutput1 )
   END_RUNG
   // the same network as SCL:
   #qOutput1 := #s260_StWtPalAbsent;
END_REGION

REGION Network 97: Transition for STATE Num:270 StWtFrTTDwnStprUp
   RUNG wire#powerrail
      Contact( #s270_StWtFrTTDwnStprUp )
      I_Contact( #sStWtResetRel )
      Contact( #sSst )
      Contact( #iStprRaise_TTDown )
      Coil( #s270_StWtFrTTDwnStprUp_T1 )
   END_RUNG
   // the same network as SCL:
   #s270_StWtFrTTDwnStprUp_T1 := #s270_StWtFrTTDwnStprUp AND NOT #sStWtResetRel AND #sSst AND #iStprRaise_TTDown;
END_REGION

REGION Network 98: STATE Num:270 StWtFrTTDwnStprUp
   RUNG wire#powerrail
      Contact( #s270_StWtFrTTDwnStprUp )
      wire#w1
      I_Contact( #sStWtResetRel )
      I_Contact( #s270_StWtFrTTDwnStprUp_T1 )
      wire#w2
      Coil( #s270_StWtFrTTDwnStprUp )
   END_RUNG
   RUNG wire#powerrail
      Contact( #s240_StWtFRTRNxtStnTTDown_T2 )
   END_RUNG wire#w1
   RUNG wire#powerrail
      Contact( #s260_StWtPalAbsent_T1 )
   END_RUNG wire#w1
   RUNG wire#w2
      { S7_GenerateENO := "TRUE" } Move(in := 270, out1 => #StateNo)
   END_RUNG
   // the same network as SCL:
   #s270_StWtFrTTDwnStprUp := (#s270_StWtFrTTDwnStprUp OR #s240_StWtFRTRNxtStnTTDown_T2 OR #s260_StWtPalAbsent_T1) AND NOT #sStWtResetRel AND NOT #s270_StWtFrTTDwnStprUp_T1;
   IF #s270_StWtFrTTDwnStprUp THEN #StateNo := 270; END_IF;
END_REGION

REGION Network 99: Actions for STATE Num:270 StWtFrTTDwnStprUp
   RUNG wire#powerrail
      Contact( #s270_StWtFrTTDwnStprUp )
      Coil( #qStprRaise_TTDown )
   END_RUNG
   // the same network as SCL:
   #qStprRaise_TTDown := #s270_StWtFrTTDwnStprUp;
END_REGION

REGION Network 100: Transition for STATE Num:280 StWtRFrOTSFRmPrev_TTUp
   RUNG wire#powerrail
      Contact( #s280_StWtRFrOTSFRmPrev_TTUp )
      I_Contact( #sStWtResetRel )
      Contact( #sSst )
      wire#w1
      Contact( #iOTS_Frm_Prev_TTUp )
      wire#w2
      Coil( #s280_StWtRFrOTSFRmPrev_TTUp_T1 )
   END_RUNG
   RUNG wire#w1
      Contact( #iPalletPrsnt_TTUp )
   END_RUNG wire#w2
   RUNG wire#w1
      Contact( #iqRx_Frm_Prev_TTUp )
   END_RUNG wire#w2
   RUNG wire#w1
      I_Contact( #iRecvAreaClr_TTUp )
   END_RUNG wire#w2
   // the same network as SCL:
   #s280_StWtRFrOTSFRmPrev_TTUp_T1 := #s280_StWtRFrOTSFRmPrev_TTUp AND NOT #sStWtResetRel AND #sSst AND (#iOTS_Frm_Prev_TTUp OR #iPalletPrsnt_TTUp OR #iqRx_Frm_Prev_TTUp OR NOT #iRecvAreaClr_TTUp);
END_REGION

REGION Network 101: STATE Num:280 StWtRFrOTSFRmPrev_TTUp
   RUNG wire#powerrail
      Contact( #s280_StWtRFrOTSFRmPrev_TTUp )
      wire#w1
      I_Contact( #sStWtResetRel )
      I_Contact( #s280_StWtRFrOTSFRmPrev_TTUp_T1 )
      wire#w2
      Coil( #s280_StWtRFrOTSFRmPrev_TTUp )
   END_RUNG
   RUNG wire#powerrail
      Contact( #s230_StWtFrTTLock_T1 )
   END_RUNG wire#w1
   RUNG wire#w2
      { S7_GenerateENO := "TRUE" } Move(in := 280, out1 => #StateNo)
   END_RUNG
   // the same network as SCL:
   #s280_StWtRFrOTSFRmPrev_TTUp := (#s280_StWtRFrOTSFRmPrev_TTUp OR #s230_StWtFrTTLock_T1) AND NOT #sStWtResetRel AND NOT #s280_StWtRFrOTSFRmPrev_TTUp_T1;
   IF #s280_StWtRFrOTSFRmPrev_TTUp THEN #StateNo := 280; END_IF;
END_REGION

REGION Network 102: Actions for STATE Num:280 StWtRFrOTSFRmPrev_TTUp
   RUNG wire#powerrail
      Contact( #s280_StWtRFrOTSFRmPrev_TTUp )
      Coil( #qRTR_Frm_TTUp )
   END_RUNG
   // the same network as SCL:
   #qRTR_Frm_TTUp := #s280_StWtRFrOTSFRmPrev_TTUp;
END_REGION

REGION Network 103: Transition for STATE Num:290 StWtFrTTUpCnvyrStrt
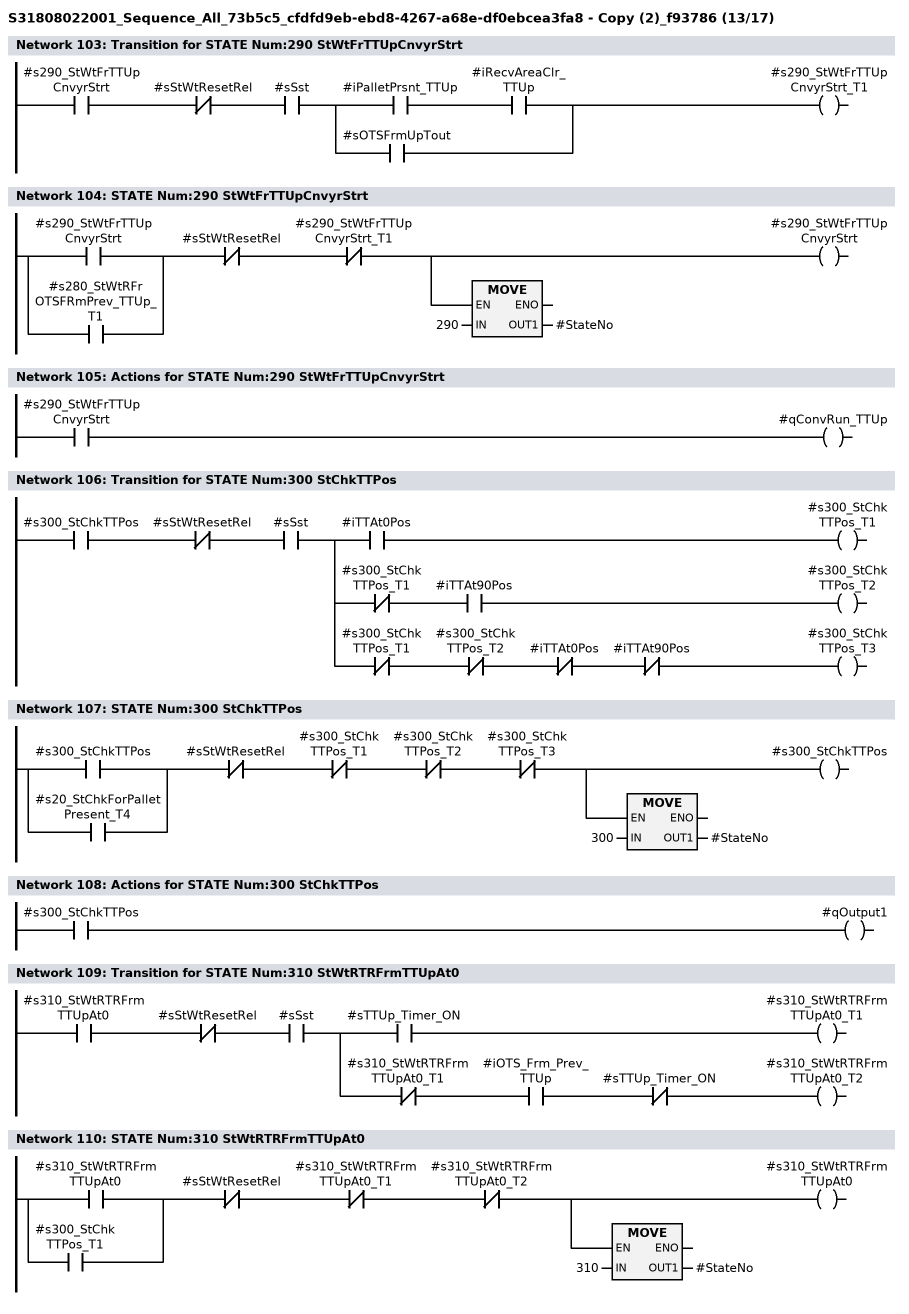
   RUNG wire#powerrail
      Contact( #s290_StWtFrTTUpCnvyrStrt )
      I_Contact( #sStWtResetRel )
      Contact( #sSst )
      wire#w1
      Contact( #iPalletPrsnt_TTUp )
      Contact( #iRecvAreaClr_TTUp )
      wire#w2
      Coil( #s290_StWtFrTTUpCnvyrStrt_T1 )
   END_RUNG
   RUNG wire#w1
      Contact( #sOTSFrmUpTout )
   END_RUNG wire#w2
   // the same network as SCL:
   #s290_StWtFrTTUpCnvyrStrt_T1 := #s290_StWtFrTTUpCnvyrStrt AND NOT #sStWtResetRel AND #sSst AND ((#iPalletPrsnt_TTUp AND #iRecvAreaClr_TTUp) OR #sOTSFrmUpTout);
END_REGION

REGION Network 104: STATE Num:290 StWtFrTTUpCnvyrStrt
   RUNG wire#powerrail
      Contact( #s290_StWtFrTTUpCnvyrStrt )
      wire#w1
      I_Contact( #sStWtResetRel )
      I_Contact( #s290_StWtFrTTUpCnvyrStrt_T1 )
      wire#w2
      Coil( #s290_StWtFrTTUpCnvyrStrt )
   END_RUNG
   RUNG wire#powerrail
      Contact( #s280_StWtRFrOTSFRmPrev_TTUp_T1 )
   END_RUNG wire#w1
   RUNG wire#w2
      { S7_GenerateENO := "TRUE" } Move(in := 290, out1 => #StateNo)
   END_RUNG
   // the same network as SCL:
   #s290_StWtFrTTUpCnvyrStrt := (#s290_StWtFrTTUpCnvyrStrt OR #s280_StWtRFrOTSFRmPrev_TTUp_T1) AND NOT #sStWtResetRel AND NOT #s290_StWtFrTTUpCnvyrStrt_T1;
   IF #s290_StWtFrTTUpCnvyrStrt THEN #StateNo := 290; END_IF;
END_REGION

REGION Network 105: Actions for STATE Num:290 StWtFrTTUpCnvyrStrt
   RUNG wire#powerrail
      Contact( #s290_StWtFrTTUpCnvyrStrt )
      Coil( #qConvRun_TTUp )
   END_RUNG
   // the same network as SCL:
   #qConvRun_TTUp := #s290_StWtFrTTUpCnvyrStrt;
END_REGION

REGION Network 106: Transition for STATE Num:300 StChkTTPos
   RUNG wire#powerrail
      Contact( #s300_StChkTTPos )
      I_Contact( #sStWtResetRel )
      Contact( #sSst )
      wire#w1
      Contact( #iTTAt0Pos )
      Coil( #s300_StChkTTPos_T1 )
   END_RUNG
   RUNG wire#w1
      I_Contact( #s300_StChkTTPos_T1 )
      Contact( #iTTAt90Pos )
      Coil( #s300_StChkTTPos_T2 )
   END_RUNG
   RUNG wire#w1
      I_Contact( #s300_StChkTTPos_T1 )
      I_Contact( #s300_StChkTTPos_T2 )
      I_Contact( #iTTAt0Pos )
      I_Contact( #iTTAt90Pos )
      Coil( #s300_StChkTTPos_T3 )
   END_RUNG
   // the same network as SCL:
   #_w1 := #s300_StChkTTPos AND NOT #sStWtResetRel AND #sSst;
   #s300_StChkTTPos_T1 := #_w1 AND #iTTAt0Pos;
   #s300_StChkTTPos_T2 := #_w1 AND NOT #s300_StChkTTPos_T1 AND #iTTAt90Pos;
   #s300_StChkTTPos_T3 := #_w1 AND NOT #s300_StChkTTPos_T1 AND NOT #s300_StChkTTPos_T2 AND NOT #iTTAt0Pos AND NOT #iTTAt90Pos;
END_REGION

REGION Network 107: STATE Num:300 StChkTTPos
   RUNG wire#powerrail
      Contact( #s300_StChkTTPos )
      wire#w1
      I_Contact( #sStWtResetRel )
      I_Contact( #s300_StChkTTPos_T1 )
      I_Contact( #s300_StChkTTPos_T2 )
      I_Contact( #s300_StChkTTPos_T3 )
      wire#w2
      Coil( #s300_StChkTTPos )
   END_RUNG
   RUNG wire#powerrail
      Contact( #s20_StChkForPalletPresent_T4 )
   END_RUNG wire#w1
   RUNG wire#w2
      { S7_GenerateENO := "TRUE" } Move(in := 300, out1 => #StateNo)
   END_RUNG
   // the same network as SCL:
   #s300_StChkTTPos := (#s300_StChkTTPos OR #s20_StChkForPalletPresent_T4) AND NOT #sStWtResetRel AND NOT #s300_StChkTTPos_T1 AND NOT #s300_StChkTTPos_T2 AND NOT #s300_StChkTTPos_T3;
   IF #s300_StChkTTPos THEN #StateNo := 300; END_IF;
END_REGION

REGION Network 108: Actions for STATE Num:300 StChkTTPos
   RUNG wire#powerrail
      Contact( #s300_StChkTTPos )
      Coil( #qOutput1 )
   END_RUNG
   // the same network as SCL:
   #qOutput1 := #s300_StChkTTPos;
END_REGION

REGION Network 109: Transition for STATE Num:310 StWtRTRFrmTTUpAt0
   RUNG wire#powerrail
      Contact( #s310_StWtRTRFrmTTUpAt0 )
      I_Contact( #sStWtResetRel )
      Contact( #sSst )
      wire#w1
      Contact( #sTTUp_Timer_ON )
      Coil( #s310_StWtRTRFrmTTUpAt0_T1 )
   END_RUNG
   RUNG wire#w1
      I_Contact( #s310_StWtRTRFrmTTUpAt0_T1 )
      Contact( #iOTS_Frm_Prev_TTUp )
      I_Contact( #sTTUp_Timer_ON )
      Coil( #s310_StWtRTRFrmTTUpAt0_T2 )
   END_RUNG
   // the same network as SCL:
   #_w1 := #s310_StWtRTRFrmTTUpAt0 AND NOT #sStWtResetRel AND #sSst;
   #s310_StWtRTRFrmTTUpAt0_T1 := #_w1 AND #sTTUp_Timer_ON;
   #s310_StWtRTRFrmTTUpAt0_T2 := #_w1 AND NOT #s310_StWtRTRFrmTTUpAt0_T1 AND #iOTS_Frm_Prev_TTUp AND NOT #sTTUp_Timer_ON;
END_REGION

REGION Network 110: STATE Num:310 StWtRTRFrmTTUpAt0
   RUNG wire#powerrail
      Contact( #s310_StWtRTRFrmTTUpAt0 )
      wire#w1
      I_Contact( #sStWtResetRel )
      I_Contact( #s310_StWtRTRFrmTTUpAt0_T1 )
      I_Contact( #s310_StWtRTRFrmTTUpAt0_T2 )
      wire#w2
      Coil( #s310_StWtRTRFrmTTUpAt0 )
   END_RUNG
   RUNG wire#powerrail
      Contact( #s300_StChkTTPos_T1 )
   END_RUNG wire#w1
   RUNG wire#w2
      { S7_GenerateENO := "TRUE" } Move(in := 310, out1 => #StateNo)
   END_RUNG
   // the same network as SCL:
   #s310_StWtRTRFrmTTUpAt0 := (#s310_StWtRTRFrmTTUpAt0 OR #s300_StChkTTPos_T1) AND NOT #sStWtResetRel AND NOT #s310_StWtRTRFrmTTUpAt0_T1 AND NOT #s310_StWtRTRFrmTTUpAt0_T2;
   IF #s310_StWtRTRFrmTTUpAt0 THEN #StateNo := 310; END_IF;
END_REGION

REGION Network 111: Actions for STATE Num:310 StWtRTRFrmTTUpAt0
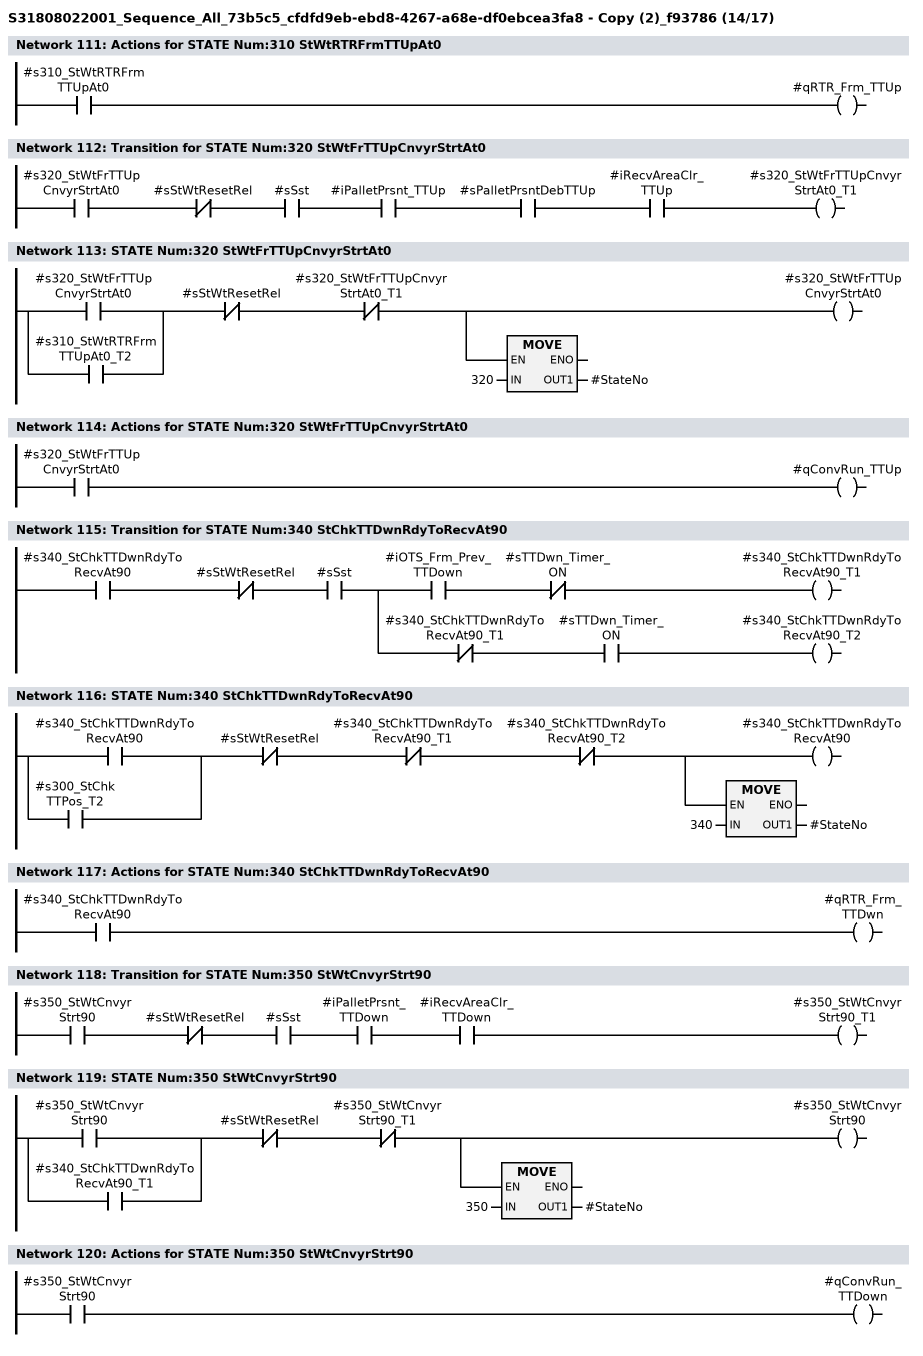
   RUNG wire#powerrail
      Contact( #s310_StWtRTRFrmTTUpAt0 )
      Coil( #qRTR_Frm_TTUp )
   END_RUNG
   // the same network as SCL:
   #qRTR_Frm_TTUp := #s310_StWtRTRFrmTTUpAt0;
END_REGION

REGION Network 112: Transition for STATE Num:320 StWtFrTTUpCnvyrStrtAt0
   RUNG wire#powerrail
      Contact( #s320_StWtFrTTUpCnvyrStrtAt0 )
      I_Contact( #sStWtResetRel )
      Contact( #sSst )
      Contact( #iPalletPrsnt_TTUp )
      Contact( #sPalletPrsntDebTTUp )
      Contact( #iRecvAreaClr_TTUp )
      Coil( #s320_StWtFrTTUpCnvyrStrtAt0_T1 )
   END_RUNG
   // the same network as SCL:
   #s320_StWtFrTTUpCnvyrStrtAt0_T1 := #s320_StWtFrTTUpCnvyrStrtAt0 AND NOT #sStWtResetRel AND #sSst AND #iPalletPrsnt_TTUp AND #sPalletPrsntDebTTUp AND #iRecvAreaClr_TTUp;
END_REGION

REGION Network 113: STATE Num:320 StWtFrTTUpCnvyrStrtAt0
   RUNG wire#powerrail
      Contact( #s320_StWtFrTTUpCnvyrStrtAt0 )
      wire#w1
      I_Contact( #sStWtResetRel )
      I_Contact( #s320_StWtFrTTUpCnvyrStrtAt0_T1 )
      wire#w2
      Coil( #s320_StWtFrTTUpCnvyrStrtAt0 )
   END_RUNG
   RUNG wire#powerrail
      Contact( #s310_StWtRTRFrmTTUpAt0_T2 )
   END_RUNG wire#w1
   RUNG wire#w2
      { S7_GenerateENO := "TRUE" } Move(in := 320, out1 => #StateNo)
   END_RUNG
   // the same network as SCL:
   #s320_StWtFrTTUpCnvyrStrtAt0 := (#s320_StWtFrTTUpCnvyrStrtAt0 OR #s310_StWtRTRFrmTTUpAt0_T2) AND NOT #sStWtResetRel AND NOT #s320_StWtFrTTUpCnvyrStrtAt0_T1;
   IF #s320_StWtFrTTUpCnvyrStrtAt0 THEN #StateNo := 320; END_IF;
END_REGION

REGION Network 114: Actions for STATE Num:320 StWtFrTTUpCnvyrStrtAt0
   RUNG wire#powerrail
      Contact( #s320_StWtFrTTUpCnvyrStrtAt0 )
      Coil( #qConvRun_TTUp )
   END_RUNG
   // the same network as SCL:
   #qConvRun_TTUp := #s320_StWtFrTTUpCnvyrStrtAt0;
END_REGION

REGION Network 115: Transition for STATE Num:340 StChkTTDwnRdyToRecvAt90
   RUNG wire#powerrail
      Contact( #s340_StChkTTDwnRdyToRecvAt90 )
      I_Contact( #sStWtResetRel )
      Contact( #sSst )
      wire#w1
      Contact( #iOTS_Frm_Prev_TTDown )
      I_Contact( #sTTDwn_Timer_ON )
      Coil( #s340_StChkTTDwnRdyToRecvAt90_T1 )
   END_RUNG
   RUNG wire#w1
      I_Contact( #s340_StChkTTDwnRdyToRecvAt90_T1 )
      Contact( #sTTDwn_Timer_ON )
      Coil( #s340_StChkTTDwnRdyToRecvAt90_T2 )
   END_RUNG
   // the same network as SCL:
   #_w1 := #s340_StChkTTDwnRdyToRecvAt90 AND NOT #sStWtResetRel AND #sSst;
   #s340_StChkTTDwnRdyToRecvAt90_T1 := #_w1 AND #iOTS_Frm_Prev_TTDown AND NOT #sTTDwn_Timer_ON;
   #s340_StChkTTDwnRdyToRecvAt90_T2 := #_w1 AND NOT #s340_StChkTTDwnRdyToRecvAt90_T1 AND #sTTDwn_Timer_ON;
END_REGION

REGION Network 116: STATE Num:340 StChkTTDwnRdyToRecvAt90
   RUNG wire#powerrail
      Contact( #s340_StChkTTDwnRdyToRecvAt90 )
      wire#w1
      I_Contact( #sStWtResetRel )
      I_Contact( #s340_StChkTTDwnRdyToRecvAt90_T1 )
      I_Contact( #s340_StChkTTDwnRdyToRecvAt90_T2 )
      wire#w2
      Coil( #s340_StChkTTDwnRdyToRecvAt90 )
   END_RUNG
   RUNG wire#powerrail
      Contact( #s300_StChkTTPos_T2 )
   END_RUNG wire#w1
   RUNG wire#w2
      { S7_GenerateENO := "TRUE" } Move(in := 340, out1 => #StateNo)
   END_RUNG
   // the same network as SCL:
   #s340_StChkTTDwnRdyToRecvAt90 := (#s340_StChkTTDwnRdyToRecvAt90 OR #s300_StChkTTPos_T2) AND NOT #sStWtResetRel AND NOT #s340_StChkTTDwnRdyToRecvAt90_T1 AND NOT #s340_StChkTTDwnRdyToRecvAt90_T2;
   IF #s340_StChkTTDwnRdyToRecvAt90 THEN #StateNo := 340; END_IF;
END_REGION

REGION Network 117: Actions for STATE Num:340 StChkTTDwnRdyToRecvAt90
   RUNG wire#powerrail
      Contact( #s340_StChkTTDwnRdyToRecvAt90 )
      Coil( #qRTR_Frm_TTDwn )
   END_RUNG
   // the same network as SCL:
   #qRTR_Frm_TTDwn := #s340_StChkTTDwnRdyToRecvAt90;
END_REGION

REGION Network 118: Transition for STATE Num:350 StWtCnvyrStrt90
   RUNG wire#powerrail
      Contact( #s350_StWtCnvyrStrt90 )
      I_Contact( #sStWtResetRel )
      Contact( #sSst )
      Contact( #iPalletPrsnt_TTDown )
      Contact( #iRecvAreaClr_TTDown )
      Coil( #s350_StWtCnvyrStrt90_T1 )
   END_RUNG
   // the same network as SCL:
   #s350_StWtCnvyrStrt90_T1 := #s350_StWtCnvyrStrt90 AND NOT #sStWtResetRel AND #sSst AND #iPalletPrsnt_TTDown AND #iRecvAreaClr_TTDown;
END_REGION

REGION Network 119: STATE Num:350 StWtCnvyrStrt90
   RUNG wire#powerrail
      Contact( #s350_StWtCnvyrStrt90 )
      wire#w1
      I_Contact( #sStWtResetRel )
      I_Contact( #s350_StWtCnvyrStrt90_T1 )
      wire#w2
      Coil( #s350_StWtCnvyrStrt90 )
   END_RUNG
   RUNG wire#powerrail
      Contact( #s340_StChkTTDwnRdyToRecvAt90_T1 )
   END_RUNG wire#w1
   RUNG wire#w2
      { S7_GenerateENO := "TRUE" } Move(in := 350, out1 => #StateNo)
   END_RUNG
   // the same network as SCL:
   #s350_StWtCnvyrStrt90 := (#s350_StWtCnvyrStrt90 OR #s340_StChkTTDwnRdyToRecvAt90_T1) AND NOT #sStWtResetRel AND NOT #s350_StWtCnvyrStrt90_T1;
   IF #s350_StWtCnvyrStrt90 THEN #StateNo := 350; END_IF;
END_REGION

REGION Network 120: Actions for STATE Num:350 StWtCnvyrStrt90
   RUNG wire#powerrail
      Contact( #s350_StWtCnvyrStrt90 )
      Coil( #qConvRun_TTDown )
   END_RUNG
   // the same network as SCL:
   #qConvRun_TTDown := #s350_StWtCnvyrStrt90;
END_REGION

REGION Network 121: Transition for STATE Num:365 StWtForTTUlkAtIbtwn
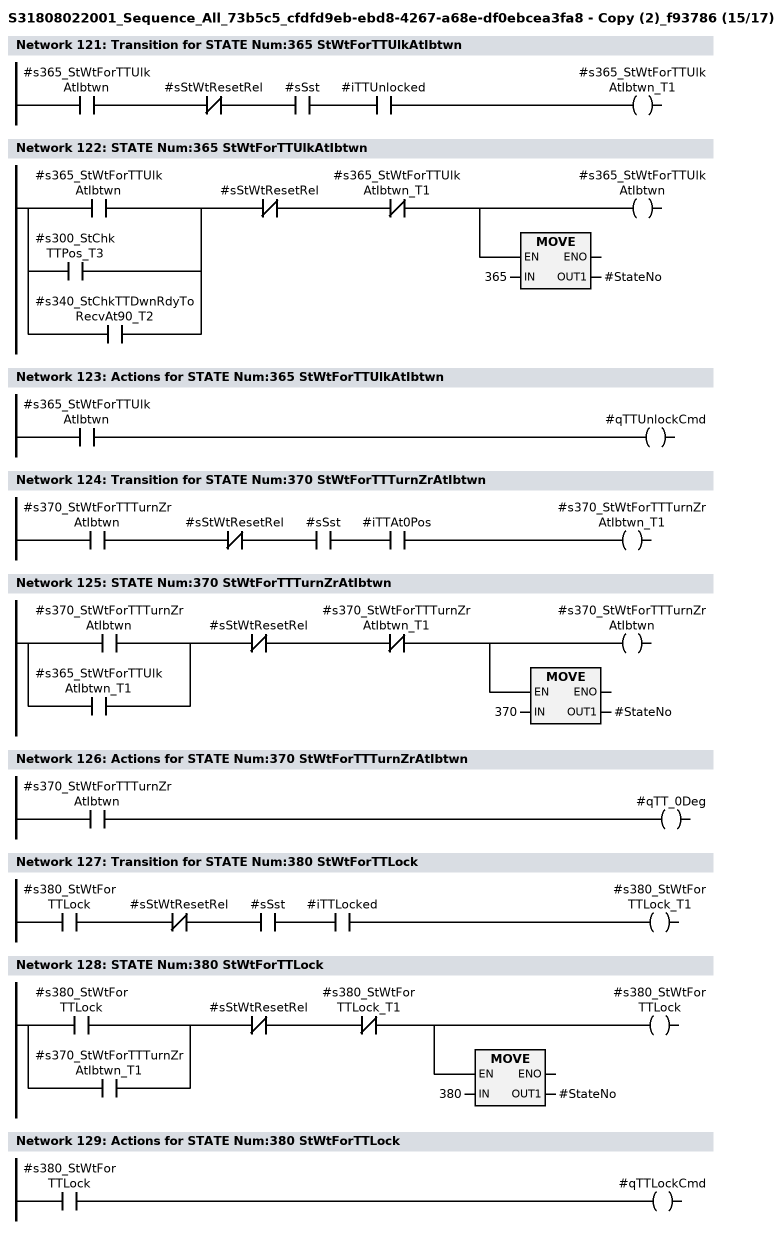
   RUNG wire#powerrail
      Contact( #s365_StWtForTTUlkAtIbtwn )
      I_Contact( #sStWtResetRel )
      Contact( #sSst )
      Contact( #iTTUnlocked )
      Coil( #s365_StWtForTTUlkAtIbtwn_T1 )
   END_RUNG
   // the same network as SCL:
   #s365_StWtForTTUlkAtIbtwn_T1 := #s365_StWtForTTUlkAtIbtwn AND NOT #sStWtResetRel AND #sSst AND #iTTUnlocked;
END_REGION

REGION Network 122: STATE Num:365 StWtForTTUlkAtIbtwn
   RUNG wire#powerrail
      Contact( #s365_StWtForTTUlkAtIbtwn )
      wire#w1
      I_Contact( #sStWtResetRel )
      I_Contact( #s365_StWtForTTUlkAtIbtwn_T1 )
      wire#w2
      Coil( #s365_StWtForTTUlkAtIbtwn )
   END_RUNG
   RUNG wire#powerrail
      Contact( #s300_StChkTTPos_T3 )
   END_RUNG wire#w1
   RUNG wire#powerrail
      Contact( #s340_StChkTTDwnRdyToRecvAt90_T2 )
   END_RUNG wire#w1
   RUNG wire#w2
      { S7_GenerateENO := "TRUE" } Move(in := 365, out1 => #StateNo)
   END_RUNG
   // the same network as SCL:
   #s365_StWtForTTUlkAtIbtwn := (#s365_StWtForTTUlkAtIbtwn OR #s300_StChkTTPos_T3 OR #s340_StChkTTDwnRdyToRecvAt90_T2) AND NOT #sStWtResetRel AND NOT #s365_StWtForTTUlkAtIbtwn_T1;
   IF #s365_StWtForTTUlkAtIbtwn THEN #StateNo := 365; END_IF;
END_REGION

REGION Network 123: Actions for STATE Num:365 StWtForTTUlkAtIbtwn
   RUNG wire#powerrail
      Contact( #s365_StWtForTTUlkAtIbtwn )
      Coil( #qTTUnlockCmd )
   END_RUNG
   // the same network as SCL:
   #qTTUnlockCmd := #s365_StWtForTTUlkAtIbtwn;
END_REGION

REGION Network 124: Transition for STATE Num:370 StWtForTTTurnZrAtIbtwn
   RUNG wire#powerrail
      Contact( #s370_StWtForTTTurnZrAtIbtwn )
      I_Contact( #sStWtResetRel )
      Contact( #sSst )
      Contact( #iTTAt0Pos )
      Coil( #s370_StWtForTTTurnZrAtIbtwn_T1 )
   END_RUNG
   // the same network as SCL:
   #s370_StWtForTTTurnZrAtIbtwn_T1 := #s370_StWtForTTTurnZrAtIbtwn AND NOT #sStWtResetRel AND #sSst AND #iTTAt0Pos;
END_REGION

REGION Network 125: STATE Num:370 StWtForTTTurnZrAtIbtwn
   RUNG wire#powerrail
      Contact( #s370_StWtForTTTurnZrAtIbtwn )
      wire#w1
      I_Contact( #sStWtResetRel )
      I_Contact( #s370_StWtForTTTurnZrAtIbtwn_T1 )
      wire#w2
      Coil( #s370_StWtForTTTurnZrAtIbtwn )
   END_RUNG
   RUNG wire#powerrail
      Contact( #s365_StWtForTTUlkAtIbtwn_T1 )
   END_RUNG wire#w1
   RUNG wire#w2
      { S7_GenerateENO := "TRUE" } Move(in := 370, out1 => #StateNo)
   END_RUNG
   // the same network as SCL:
   #s370_StWtForTTTurnZrAtIbtwn := (#s370_StWtForTTTurnZrAtIbtwn OR #s365_StWtForTTUlkAtIbtwn_T1) AND NOT #sStWtResetRel AND NOT #s370_StWtForTTTurnZrAtIbtwn_T1;
   IF #s370_StWtForTTTurnZrAtIbtwn THEN #StateNo := 370; END_IF;
END_REGION

REGION Network 126: Actions for STATE Num:370 StWtForTTTurnZrAtIbtwn
   RUNG wire#powerrail
      Contact( #s370_StWtForTTTurnZrAtIbtwn )
      Coil( #qTT_0Deg )
   END_RUNG
   // the same network as SCL:
   #qTT_0Deg := #s370_StWtForTTTurnZrAtIbtwn;
END_REGION

REGION Network 127: Transition for STATE Num:380 StWtForTTLock
   RUNG wire#powerrail
      Contact( #s380_StWtForTTLock )
      I_Contact( #sStWtResetRel )
      Contact( #sSst )
      Contact( #iTTLocked )
      Coil( #s380_StWtForTTLock_T1 )
   END_RUNG
   // the same network as SCL:
   #s380_StWtForTTLock_T1 := #s380_StWtForTTLock AND NOT #sStWtResetRel AND #sSst AND #iTTLocked;
END_REGION

REGION Network 128: STATE Num:380 StWtForTTLock
   RUNG wire#powerrail
      Contact( #s380_StWtForTTLock )
      wire#w1
      I_Contact( #sStWtResetRel )
      I_Contact( #s380_StWtForTTLock_T1 )
      wire#w2
      Coil( #s380_StWtForTTLock )
   END_RUNG
   RUNG wire#powerrail
      Contact( #s370_StWtForTTTurnZrAtIbtwn_T1 )
   END_RUNG wire#w1
   RUNG wire#w2
      { S7_GenerateENO := "TRUE" } Move(in := 380, out1 => #StateNo)
   END_RUNG
   // the same network as SCL:
   #s380_StWtForTTLock := (#s380_StWtForTTLock OR #s370_StWtForTTTurnZrAtIbtwn_T1) AND NOT #sStWtResetRel AND NOT #s380_StWtForTTLock_T1;
   IF #s380_StWtForTTLock THEN #StateNo := 380; END_IF;
END_REGION

REGION Network 129: Actions for STATE Num:380 StWtForTTLock
   RUNG wire#powerrail
      Contact( #s380_StWtForTTLock )
      Coil( #qTTLockCmd )
   END_RUNG
   // the same network as SCL:
   #qTTLockCmd := #s380_StWtForTTLock;
END_REGION

REGION Network 130: Condition1 for STATE Num:400 Wait for all 2 Sub Sequences to complete
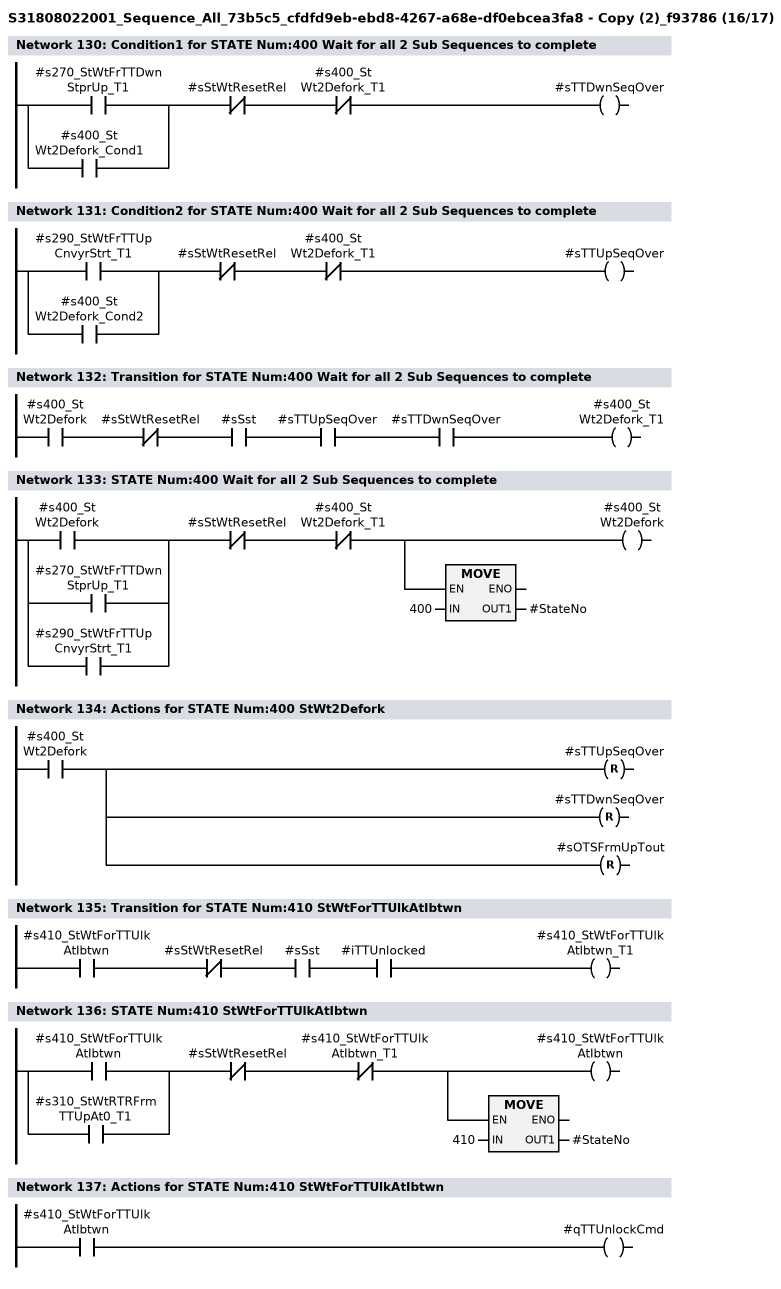
   RUNG wire#powerrail
      Contact( #s270_StWtFrTTDwnStprUp_T1 )
      wire#w1
      I_Contact( #sStWtResetRel )
      I_Contact( #s400_StWt2Defork_T1 )
      Coil( #sTTDwnSeqOver )
   END_RUNG
   RUNG wire#powerrail
      Contact( #s400_StWt2Defork_Cond1 )
   END_RUNG wire#w1
   // the same network as SCL:
   #sTTDwnSeqOver := (#s270_StWtFrTTDwnStprUp_T1 OR #s400_StWt2Defork_Cond1) AND NOT #sStWtResetRel AND NOT #s400_StWt2Defork_T1;
END_REGION

REGION Network 131: Condition2 for STATE Num:400 Wait for all 2 Sub Sequences to complete
   RUNG wire#powerrail
      Contact( #s290_StWtFrTTUpCnvyrStrt_T1 )
      wire#w1
      I_Contact( #sStWtResetRel )
      I_Contact( #s400_StWt2Defork_T1 )
      Coil( #sTTUpSeqOver )
   END_RUNG
   RUNG wire#powerrail
      Contact( #s400_StWt2Defork_Cond2 )
   END_RUNG wire#w1
   // the same network as SCL:
   #sTTUpSeqOver := (#s290_StWtFrTTUpCnvyrStrt_T1 OR #s400_StWt2Defork_Cond2) AND NOT #sStWtResetRel AND NOT #s400_StWt2Defork_T1;
END_REGION

REGION Network 132: Transition for STATE Num:400 Wait for all 2 Sub Sequences to complete
   RUNG wire#powerrail
      Contact( #s400_StWt2Defork )
      I_Contact( #sStWtResetRel )
      Contact( #sSst )
      Contact( #sTTUpSeqOver )
      Contact( #sTTDwnSeqOver )
      Coil( #s400_StWt2Defork_T1 )
   END_RUNG
   // the same network as SCL:
   #s400_StWt2Defork_T1 := #s400_StWt2Defork AND NOT #sStWtResetRel AND #sSst AND #sTTUpSeqOver AND #sTTDwnSeqOver;
END_REGION

REGION Network 133: STATE Num:400 Wait for all 2 Sub Sequences to complete
   RUNG wire#powerrail
      Contact( #s400_StWt2Defork )
      wire#w1
      I_Contact( #sStWtResetRel )
      I_Contact( #s400_StWt2Defork_T1 )
      wire#w2
      Coil( #s400_StWt2Defork )
   END_RUNG
   RUNG wire#powerrail
      Contact( #s270_StWtFrTTDwnStprUp_T1 )
   END_RUNG wire#w1
   RUNG wire#powerrail
      Contact( #s290_StWtFrTTUpCnvyrStrt_T1 )
   END_RUNG wire#w1
   RUNG wire#w2
      { S7_GenerateENO := "TRUE" } Move(in := 400, out1 => #StateNo)
   END_RUNG
   // the same network as SCL:
   #s400_StWt2Defork := (#s400_StWt2Defork OR #s270_StWtFrTTDwnStprUp_T1 OR #s290_StWtFrTTUpCnvyrStrt_T1) AND NOT #sStWtResetRel AND NOT #s400_StWt2Defork_T1;
   IF #s400_StWt2Defork THEN #StateNo := 400; END_IF;
END_REGION

REGION Network 134: Actions for STATE Num:400 StWt2Defork
   RUNG wire#powerrail
      Contact( #s400_StWt2Defork )
      wire#w1
      R_Coil( #sTTUpSeqOver )
   END_RUNG
   RUNG wire#w1
      R_Coil( #sTTDwnSeqOver )
   END_RUNG
   RUNG wire#w1
      R_Coil( #sOTSFrmUpTout )
   END_RUNG
   // the same network as SCL:
   IF #s400_StWt2Defork THEN
       #sTTUpSeqOver := FALSE;
       #sTTDwnSeqOver := FALSE;
       #sOTSFrmUpTout := FALSE;
   END_IF;
END_REGION

REGION Network 135: Transition for STATE Num:410 StWtForTTUlkAtIbtwn
   RUNG wire#powerrail
      Contact( #s410_StWtForTTUlkAtIbtwn )
      I_Contact( #sStWtResetRel )
      Contact( #sSst )
      Contact( #iTTUnlocked )
      Coil( #s410_StWtForTTUlkAtIbtwn_T1 )
   END_RUNG
   // the same network as SCL:
   #s410_StWtForTTUlkAtIbtwn_T1 := #s410_StWtForTTUlkAtIbtwn AND NOT #sStWtResetRel AND #sSst AND #iTTUnlocked;
END_REGION

REGION Network 136: STATE Num:410 StWtForTTUlkAtIbtwn
   RUNG wire#powerrail
      Contact( #s410_StWtForTTUlkAtIbtwn )
      wire#w1
      I_Contact( #sStWtResetRel )
      I_Contact( #s410_StWtForTTUlkAtIbtwn_T1 )
      wire#w2
      Coil( #s410_StWtForTTUlkAtIbtwn )
   END_RUNG
   RUNG wire#powerrail
      Contact( #s310_StWtRTRFrmTTUpAt0_T1 )
   END_RUNG wire#w1
   RUNG wire#w2
      { S7_GenerateENO := "TRUE" } Move(in := 410, out1 => #StateNo)
   END_RUNG
   // the same network as SCL:
   #s410_StWtForTTUlkAtIbtwn := (#s410_StWtForTTUlkAtIbtwn OR #s310_StWtRTRFrmTTUpAt0_T1) AND NOT #sStWtResetRel AND NOT #s410_StWtForTTUlkAtIbtwn_T1;
   IF #s410_StWtForTTUlkAtIbtwn THEN #StateNo := 410; END_IF;
END_REGION

REGION Network 137: Actions for STATE Num:410 StWtForTTUlkAtIbtwn
   RUNG wire#powerrail
      Contact( #s410_StWtForTTUlkAtIbtwn )
      Coil( #qTTUnlockCmd )
   END_RUNG
   // the same network as SCL:
   #qTTUnlockCmd := #s410_StWtForTTUlkAtIbtwn;
END_REGION

REGION Network 138: Transition for STATE Num:415 StWtForTTTurn90AtIbtwn
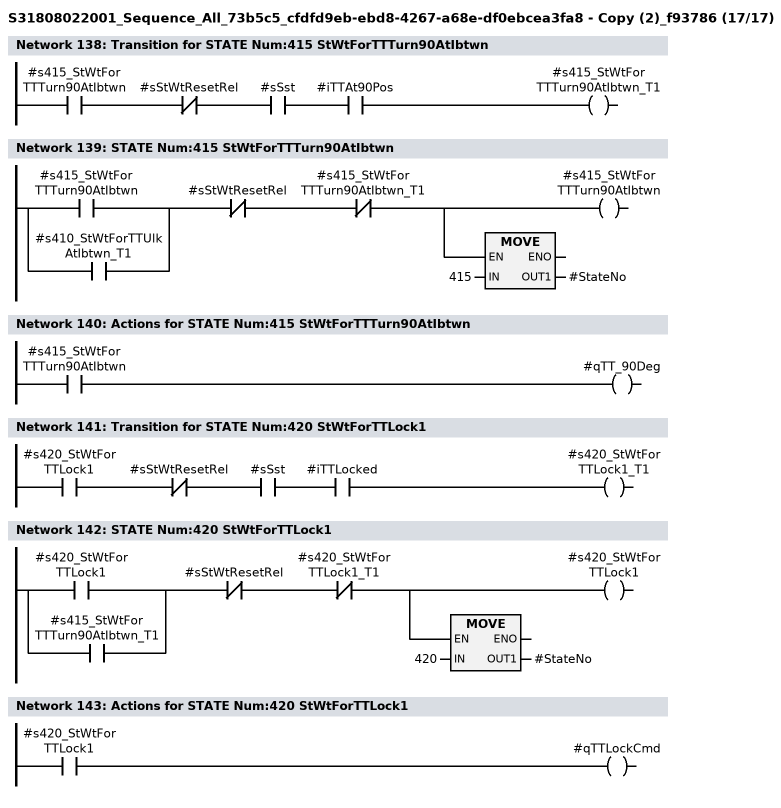
   RUNG wire#powerrail
      Contact( #s415_StWtForTTTurn90AtIbtwn )
      I_Contact( #sStWtResetRel )
      Contact( #sSst )
      Contact( #iTTAt90Pos )
      Coil( #s415_StWtForTTTurn90AtIbtwn_T1 )
   END_RUNG
   // the same network as SCL:
   #s415_StWtForTTTurn90AtIbtwn_T1 := #s415_StWtForTTTurn90AtIbtwn AND NOT #sStWtResetRel AND #sSst AND #iTTAt90Pos;
END_REGION

REGION Network 139: STATE Num:415 StWtForTTTurn90AtIbtwn
   RUNG wire#powerrail
      Contact( #s415_StWtForTTTurn90AtIbtwn )
      wire#w1
      I_Contact( #sStWtResetRel )
      I_Contact( #s415_StWtForTTTurn90AtIbtwn_T1 )
      wire#w2
      Coil( #s415_StWtForTTTurn90AtIbtwn )
   END_RUNG
   RUNG wire#powerrail
      Contact( #s410_StWtForTTUlkAtIbtwn_T1 )
   END_RUNG wire#w1
   RUNG wire#w2
      { S7_GenerateENO := "TRUE" } Move(in := 415, out1 => #StateNo)
   END_RUNG
   // the same network as SCL:
   #s415_StWtForTTTurn90AtIbtwn := (#s415_StWtForTTTurn90AtIbtwn OR #s410_StWtForTTUlkAtIbtwn_T1) AND NOT #sStWtResetRel AND NOT #s415_StWtForTTTurn90AtIbtwn_T1;
   IF #s415_StWtForTTTurn90AtIbtwn THEN #StateNo := 415; END_IF;
END_REGION

REGION Network 140: Actions for STATE Num:415 StWtForTTTurn90AtIbtwn
   RUNG wire#powerrail
      Contact( #s415_StWtForTTTurn90AtIbtwn )
      Coil( #qTT_90Deg )
   END_RUNG
   // the same network as SCL:
   #qTT_90Deg := #s415_StWtForTTTurn90AtIbtwn;
END_REGION

REGION Network 141: Transition for STATE Num:420 StWtForTTLock1
   RUNG wire#powerrail
      Contact( #s420_StWtForTTLock1 )
      I_Contact( #sStWtResetRel )
      Contact( #sSst )
      Contact( #iTTLocked )
      Coil( #s420_StWtForTTLock1_T1 )
   END_RUNG
   // the same network as SCL:
   #s420_StWtForTTLock1_T1 := #s420_StWtForTTLock1 AND NOT #sStWtResetRel AND #sSst AND #iTTLocked;
END_REGION

REGION Network 142: STATE Num:420 StWtForTTLock1
   RUNG wire#powerrail
      Contact( #s420_StWtForTTLock1 )
      wire#w1
      I_Contact( #sStWtResetRel )
      I_Contact( #s420_StWtForTTLock1_T1 )
      wire#w2
      Coil( #s420_StWtForTTLock1 )
   END_RUNG
   RUNG wire#powerrail
      Contact( #s415_StWtForTTTurn90AtIbtwn_T1 )
   END_RUNG wire#w1
   RUNG wire#w2
      { S7_GenerateENO := "TRUE" } Move(in := 420, out1 => #StateNo)
   END_RUNG
   // the same network as SCL:
   #s420_StWtForTTLock1 := (#s420_StWtForTTLock1 OR #s415_StWtForTTTurn90AtIbtwn_T1) AND NOT #sStWtResetRel AND NOT #s420_StWtForTTLock1_T1;
   IF #s420_StWtForTTLock1 THEN #StateNo := 420; END_IF;
END_REGION

REGION Network 143: Actions for STATE Num:420 StWtForTTLock1
   RUNG wire#powerrail
      Contact( #s420_StWtForTTLock1 )
      Coil( #qTTLockCmd )
   END_RUNG
   // the same network as SCL:
   #qTTLockCmd := #s420_StWtForTTLock1;
END_REGION
END_FUNCTION_BLOCK
